        MoveJ speed 60 deg/s, acceleration 80 deg/s^2 (useActiveTCP=true optimoveEnabled=false optiMoveSpeed=0.3 optiMoveAcceleration=0.09) feature=Base
          Waypoint Waypoint_104: TCP in base x=-333.293 y=-480.744 z=350.142 mm, rx=2.2175 ry=0.1409 rz=2.2091 rad; joints [-82.414, -101.687, -97.87, -162.913, 4.302, 96.426] deg
        SuppressedNode
          Weight_value := get_weight()
    SuppressedNode
      Case (caseValue=38)
        SuppressedNode
          URCap VISOR Robotic App (SensoPart VISOR Robotic, SensoPart Industriesensorik GmbH) dataModel(visorAppTemplate=1); state(isChildrenLocked=true)
            URCap Easy Pick Setup (SensoPart VISOR Robotic, SensoPart Industriesensorik GmbH) dataModel(visorId=0, visorSetJob=true, visorJobName=Container_S_rack, visorImageAcqSetup=2, visorSetupStatus=2); state(isChildrenLocked=true)
            URCap Process (SensoPart VISOR Robotic, SensoPart Industriesensorik GmbH) dataModel(Variable(key=visorCounterVar, variable(name=easyPickCount_4, initializeExpression=0)), Variable(key=visorPartsFoundVar, variable(name=easyPickParts_4, initializeExpression=0))); state(isChildrenLocked=true)
              URCap Image Acquisition Pose (SensoPart VISOR Robotic, SensoPart Industriesensorik GmbH) state(isChildrenLocked=true)
              URCap Object Detected (SensoPart VISOR Robotic, SensoPart Industriesensorik GmbH) state(isChildrenLocked=true)
                Folder Open Gripper
                  Placeholder
                URCap Approach Pose (SensoPart VISOR Robotic, SensoPart Industriesensorik GmbH) state(isChildrenLocked=true)
                URCap Target Pose (SensoPart VISOR Robotic, SensoPart Industriesensorik GmbH) state(isChildrenLocked=true)
                Folder Close Gripper
                  Placeholder
                URCap Exit Pose (SensoPart VISOR Robotic, SensoPart Industriesensorik GmbH) state(isChildrenLocked=true)
              URCap No Object Detected (SensoPart VISOR Robotic, SensoPart Industriesensorik GmbH) dataModel(Variable(key=visorNoObjCountVar, variable(name=easyPickNoObj_4, initializeExpression=0)))
                Placeholder
    Case (caseValue=39)
      Folder Powder container Pick [hidden by the author, left out]
    Case (caseValue=40)
      Folder Decap Container  [hidden by the author, left out]
    Case (caseValue=41)
      Folder Place the open PowderA container & dosing
        SuppressedNode
          Script: tilt_to_home()
        SuppressedNode
          Script: tilt_send(4)
        URCap VISOR Robotic App (SensoPart VISOR Robotic, SensoPart Industriesensorik GmbH) dataModel(visorAppTemplate=1); state(isChildrenLocked=true)
          URCap Easy Pick Setup (SensoPart VISOR Robotic, SensoPart Industriesensorik GmbH) dataModel(visorId=0, visorImageAcqSetup=2, visorDetector=1, visorSetJob=true, visorOffsetSet=true, visorImageAcqSource=2, visorJobName=PoTS, visorSetupStatus=3, Pose(key=visorGripPose, Position(key=posePosition, Length(key=X value=-0.729991 unit=M), Length(key=Y value=-0.185228 unit=M), Length(key=Z value=0.248335 unit=M)), Rotation(key=poseRotation, Angle(key=RX value=-0.919003 unit=RAD), Angle(key=RY value=1.612625 unit=RAD), Angle(key=RZ value=-1.647622 unit=RAD))), Feature(key=visorImageAcqFeature name=Trigger)); state(isChildrenLocked=true)
          URCap Process (SensoPart VISOR Robotic, SensoPart Industriesensorik GmbH) dataModel(Variable(key=visorCounterVar, variable(name=easyPickCount_7, initializeExpression=0)), Variable(key=visorPartsFoundVar, variable(name=easyPickParts_7, initializeExpression=0))); state(isChildrenLocked=true)
            URCap Image Acquisition Pose (SensoPart VISOR Robotic, SensoPart Industriesensorik GmbH) state(isChildrenLocked=true)
            URCap Object Detected (SensoPart VISOR Robotic, SensoPart Industriesensorik GmbH) state(isChildrenLocked=true)
              Folder Open Gripper
                URCap Gripper (Robotiq_Grippers, Robotiq Inc.) dataModel(position=0.0, force=30.19607843137255, speed=30.19607843137255, positionInDouble=0.0, forceInDouble=30.19607843137255, speedInDouble=30.19607843137255, slaveIds=[9], blocking=true)
                SuppressedNode
                  Set NoAction tcp=TCP_fingers
                SuppressedNode
                  Wait Sleep waitTime=0.2
                MoveL speed 250 mm/s, acceleration 1200 mm/s^2 (useActiveTCP=true optimoveEnabled=false optiMoveSpeed=0.3 optiMoveAcceleration=0.09) feature=Base
                  Waypoint OP_PowderA2: TCP in base x=9.371 y=-409.434 z=294.169 mm, rx=-0.8233 ry=1.7094 rz=-1.6983 rad; joints [-57.265, -122.586, -76.992, -161.25, 72.295, 1.124] deg; TCP offset x=0 y=0 z=161 mm, rx=3.1415 ry=0 rz=0 rad
                  Waypoint OP_PowderA_ab_1: TCP in base x=-12.145 y=-363.335 z=315.326 mm, rx=-0.7771 ry=1.753 rz=-1.7409 rad; joints [-58.232, -116.012, -83.989, -160.83, 75.01, 1.147] deg; TCP offset x=0 y=0 z=161 mm, rx=3.1415 ry=0 rz=0 rad
                  Waypoint OP_PowderA_pick: TCP in base x=-19.99 y=-367.909 z=180.101 mm, rx=-0.5462 ry=1.936 rz=-1.9301 rad; joints [-66.516, -128.259, -85.768, -146.461, 83.267, 1.188] deg
                  URCap Gripper (Robotiq_Grippers, Robotiq Inc.) dataModel(position=100.0, force=30.19607843137255, speed=30.19607843137255, positionInDouble=100.0, forceInDouble=30.19607843137255, speedInDouble=30.19607843137255, slaveIds=[9], blocking=true)
                  Wait Sleep waitTime=0.5
                  Set DigitalOutput pin=GRP_3F_Open; digitalValue=1
                  SuppressedNode
                    Script: Motors_off()
                  Waypoint OP_PowderA_ab_2: motionParameters(jointSpeed=1.047198 jointAcceleration=1.396263 cartesianSpeed=0.05 cartesianAcceleration=0.3); TCP in base x=-12.145 y=-363.335 z=315.326 mm, rx=-0.7771 ry=1.753 rz=-1.7409 rad; joints [-58.232, -116.012, -83.989, -160.83, 75.01, 1.147] deg
                  Waypoint Op_PowA_wP: TCP in base x=-173.728 y=-372.934 z=295.117 mm, rx=-0.9724 ry=1.541 rz=-1.5487 rad; joints [-67.269, -106.894, -99.849, -153.52, 49.211, 1.028] deg
              URCap Approach Pose (SensoPart VISOR Robotic, SensoPart Industriesensorik GmbH) dataModel(visorOffsetZ=0.0, visorJointSpeed=25.0, visorJointAcc=30.0); state(isChildrenLocked=true)
              URCap Target Pose (SensoPart VISOR Robotic, SensoPart Industriesensorik GmbH) dataModel(visorToolSpeed=50.0, visorToolAcc=100.0); state(isChildrenLocked=true)
              Folder Close Gripper
                container_place := get_actual_tcp_pose()
                SuppressedNode
                  radius := 0.035
                SuppressedNode
                  PoTS_place_abov := pose_trans(container_place, p[0,0,radius,0,0,0])
                SuppressedNode
                  MoveL speed 50 mm/s, acceleration 500 mm/s^2 (useActiveTCP=true optimoveEnabled=false optiMoveSpeed=0.3 optiMoveAcceleration=0.09) feature=Base
                    Waypoint Variable (Variable): variable(name=PoTS_place_abov)
                target_pose := pose_trans(container_place, p[0,0.09,0,0,0,0])
                MoveL speed 50 mm/s, acceleration 500 mm/s^2 (useActiveTCP=true optimoveEnabled=false optiMoveSpeed=0.3 optiMoveAcceleration=0.09) feature=Base
                  Waypoint Variable (Variable): motionParameters(jointSpeed=1.047198 jointAcceleration=1.396263 cartesianSpeed=0.05 cartesianAcceleration=0.3); variable=target_pose
                URCap Gripper (Robotiq_Grippers, Robotiq Inc.) dataModel(position=0.0, force=30.19607843137255, speed=30.19607843137255, positionInDouble=0.0, forceInDouble=30.19607843137255, speedInDouble=30.19607843137255, slaveIds=[9], blocking=true)
              URCap Exit Pose (SensoPart VISOR Robotic, SensoPart Industriesensorik GmbH) dataModel(visorOffsetZ=-50.0); state(isChildrenLocked=true)
            URCap No Object Detected (SensoPart VISOR Robotic, SensoPart Industriesensorik GmbH) dataModel(Variable(key=visorNoObjCountVar, variable(name=easyPickNoObj_7, initializeExpression=0)))
              Popup Message (haltProgram=false message=No weigh scale detected inputType=Text)
        place_pose := get_actual_tcp_pose()
        Script: center_pose()
        SuppressedNode
          center_tilt_pos := P_center
        MoveJ speed 60 deg/s, acceleration 80 deg/s^2 (useActiveTCP=true optimoveEnabled=false optiMoveSpeed=0.3 optiMoveAcceleration=0.09) feature=Base
          Waypoint Waypoint_1: TCP in base x=-451.049 y=-340.589 z=308.224 mm, rx=0.0971 ry=0.091 rz=-1.5784 rad; joints [-127.334, -100.578, -80.109, -94.907, 86.186, -126.663] deg
    Case (caseValue=42)
      Folder Powder Emptying [hidden by the author, left out]
    Case (caseValue=43)
      Folder Powder dosing
        SuppressedNode
          Script: zero_scale()
        Script: send_target_info()
        Script: send_powder_info()
        switch_spat_M := True
        switch_spat_S := True
        switch_spat_F_S := True
        Timer (action=Start) variable(name=Dosing_time)
        SuppressedNode
          Script: tilt_to_home()
        SuppressedNode
          Folder spatula_selection test
            weight_value := get_weight()
            diff := target_weight-weight_value
            Script: scooping_init()
            Script: compute_level_percent(W_now, weight_value)
            Script: spatula = select_spatula(Pow_name, level, diff)
        URCap VISOR Robotic App (SensoPart VISOR Robotic, SensoPart Industriesensorik GmbH) dataModel(visorAppTemplate=1); state(isChildrenLocked=true)
          URCap Easy Pick Setup (SensoPart VISOR Robotic, SensoPart Industriesensorik GmbH) dataModel(visorId=0, visorSetJob=true, visorImageAcqSetup=2, visorCalibSetNo=9, visorDetector=1, visorImageAcqSource=2, visorJobName=Weight_scale, visorOffsetSet=true, visorSetupStatus=3, Pose(key=visorGripPose, Position(key=posePosition, Length(key=X value=-0.45122 unit=M), Length(key=Y value=0.110677 unit=M), Length(key=Z value=0.129785 unit=M)), Rotation(key=poseRotation, Angle(key=RX value=0.852924 unit=RAD), Angle(key=RY value=1.33496 unit=RAD), Angle(key=RZ value=-0.958582 unit=RAD))), Feature(key=visorImageAcqFeature name=Trigger)); state(isChildrenLocked=true)
          URCap Process (SensoPart VISOR Robotic, SensoPart Industriesensorik GmbH) dataModel(Variable(key=visorCounterVar, variable=easyPickCount_4), Variable(key=visorPartsFoundVar, variable=easyPickParts_4)); state(isChildrenLocked=true)
            URCap Image Acquisition Pose (SensoPart VISOR Robotic, SensoPart Industriesensorik GmbH) state(isChildrenLocked=true)
            URCap Object Detected (SensoPart VISOR Robotic, SensoPart Industriesensorik GmbH) state(isChildrenLocked=true)
              Folder Open Gripper
                Script: tare_scale()
                Wait Sleep waitTime=0.2
                weight_value := get_weight()
                Wait Sleep waitTime=0.2
                diff := target_weight-weight_value
                Script: scooping_init()
                Script: compute_level_percent(W_now, weight_value)
                Script: send_level_info()
                spatula := select_spatula(Pow_name, level, diff)
                SuppressedNode
                  spatula := select_spatula(Flowability,level,diff,density)
                SuppressedNode
                  Script: spatula = "spatula_M"
                Wait Sleep waitTime=0.2
                Script: send_spatula_info()
                If spatula ≟ "spatula_L"
                  MoveJ speed 60 deg/s, acceleration 80 deg/s^2 (useActiveTCP=true optimoveEnabled=false optiMoveSpeed=0.3 optiMoveAcceleration=0.09) feature=Base
                    Waypoint Spatula_otw: TCP in base x=-222.06 y=-318.141 z=425.288 mm, rx=-0.0004 ry=-0.0001 rz=3.0344 rad; joints [-104.723, -74.795, -88.594, -106.601, 90.132, -8.655] deg
                    Waypoint pick_spat_L_abv: TCP in base x=239.059 y=-67.213 z=280.721 mm, rx=0 ry=-0.0005 rz=3.1068 rad; joints [16.774, -49.077, -122.624, -98.282, 90.162, 108.776] deg
                  MoveL speed 250 mm/s, acceleration 1200 mm/s^2 (useActiveTCP=true optimoveEnabled=false optiMoveSpeed=0.3 optiMoveAcceleration=0.09) feature=Base
                    Waypoint spat_L_pick: TCP in base x=242.469 y=-67.302 z=193.171 mm, rx=0 ry=-0.0005 rz=3.1068 rad; joints [16.429, -49.275, -135.385, -85.324, 90.17, 108.483] deg
                    URCap Gripper (Robotiq_Grippers, Robotiq Inc.) dataModel(position=100.0, force=30.0, speed=0.0, positionInDouble=100.0, forceInDouble=30.0, speedInDouble=0.0, slaveIds=[9], blocking=true)
                    Waypoint spat_L_lift: motionParameters(blendRadius=0.01); TCP in base x=245.402 y=-67.432 z=289.049 mm, rx=0 ry=-0.0005 rz=3.1068 rad; joints [16.24, -50.411, -121.005, -98.568, 90.16, 108.238] deg
                    Waypoint spat_L_side: motionParameters(blendRadius=0.01); TCP in base x=247.134 y=-17.634 z=289.063 mm, rx=0 ry=-0.0005 rz=3.1068 rad; joints [28.487, -49.174, -121.365, -99.443, 90.16, 120.484] deg
                    Waypoint spat_L_up: motionParameters(blendRadius=0.05); TCP in base x=247.136 y=-17.665 z=397.131 mm, rx=0 ry=-0.0005 rz=3.1068 rad; joints [28.565, -53.55, -103.607, -112.824, 90.132, 120.503] deg
                  MoveJ speed 60 deg/s, acceleration 80 deg/s^2 (useActiveTCP=true optimoveEnabled=false optiMoveSpeed=0.3 optiMoveAcceleration=0.09) feature=Base
                    Waypoint Spatula_otw: TCP in base x=-222.06 y=-318.141 z=425.288 mm, rx=-0.0004 ry=-0.0001 rz=3.0344 rad; joints [-104.723, -74.795, -88.594, -106.601, 90.132, -8.655] deg
                ElseIf spatula ≟"spatula_M"
                  MoveJ speed 60 deg/s, acceleration 80 deg/s^2 (useActiveTCP=true optimoveEnabled=false optiMoveSpeed=0.3 optiMoveAcceleration=0.09) feature=Base
                    Waypoint Spatula_otw: TCP in base x=-222.06 y=-318.141 z=425.288 mm, rx=-0.0004 ry=-0.0001 rz=3.0344 rad; joints [-104.723, -74.795, -88.594, -106.601, 90.132, -8.655] deg
                    Waypoint spat_M_up: motionParameters(blendRadius=0.05); TCP in base x=245.496 y=-112.113 z=420.344 mm, rx=0 ry=-0.0005 rz=3.0677 rad; joints [5.167, -58.065, -98.393, -113.528, 90.127, 99.337] deg
                  MoveL speed 250 mm/s, acceleration 1200 mm/s^2 (useActiveTCP=true optimoveEnabled=false optiMoveSpeed=0.3 optiMoveAcceleration=0.09) feature=Base
                    Waypoint spat_M_pick: TCP in base x=244.674 y=-111.985 z=192.299 mm, rx=0 ry=-0.0005 rz=3.0677 rad; joints [5.062, -53.127, -134.29, -82.569, 90.166, 99.363] deg
                    URCap Gripper (Robotiq_Grippers, Robotiq Inc.) dataModel(position=100.0, force=30.0, speed=0.0, positionInDouble=100.0, forceInDouble=30.0, speedInDouble=0.0, slaveIds=[9], blocking=true)
                    Waypoint spat_M_up: motionParameters(blendRadius=0.05); TCP in base x=245.496 y=-112.113 z=420.344 mm, rx=0 ry=-0.0005 rz=3.0677 rad; joints [5.167, -58.065, -98.393, -113.528, 90.127, 99.337] deg
                    Waypoint Spatula_otw: TCP in base x=-222.06 y=-318.141 z=425.288 mm, rx=-0.0004 ry=-0.0001 rz=3.0344 rad; joints [-104.723, -74.795, -88.594, -106.601, 90.132, -8.655] deg
                  switch_spat_M := False
                ElseIf spatula≟"spatula_S"
                  MoveJ speed 60 deg/s, acceleration 80 deg/s^2 (useActiveTCP=true optimoveEnabled=false optiMoveSpeed=0.3 optiMoveAcceleration=0.09) feature=Base
                    Waypoint Spatula_otw: TCP in base x=-222.06 y=-318.141 z=425.288 mm, rx=-0.0004 ry=-0.0001 rz=3.0344 rad; joints [-104.723, -74.795, -88.594, -106.601, 90.132, -8.655] deg
                    Waypoint spat_S_Up_7: motionParameters(blendRadius=0.05); TCP in base x=252.088 y=-159.242 z=423.282 mm, rx=0 ry=-0.0005 rz=3.0677 rad; joints [-5.618, -62.24, -96.192, -111.556, 90.127, 88.551] deg
                  MoveL speed 250 mm/s, acceleration 1200 mm/s^2 (useActiveTCP=true optimoveEnabled=false optiMoveSpeed=0.3 optiMoveAcceleration=0.09) feature=Base
                    Waypoint spat_S_Pick_4: TCP in base x=245.377 y=-158.668 z=192.286 mm, rx=0 ry=-0.0005 rz=3.0677 rad; joints [-5.78, -57.937, -132.467, -79.585, 90.161, 88.525] deg
                    URCap Gripper (Robotiq_Grippers, Robotiq Inc.) dataModel(position=100.0, force=30.0, speed=0.0, positionInDouble=100.0, forceInDouble=30.0, speedInDouble=0.0, slaveIds=[9], blocking=true)
                    Waypoint spat_S_Up_8: motionParameters(blendRadius=0.05); TCP in base x=252.088 y=-159.242 z=423.282 mm, rx=0 ry=-0.0005 rz=3.0677 rad; joints [-5.618, -62.24, -96.192, -111.556, 90.127, 88.551] deg
                    Waypoint Spatula_otw: TCP in base x=-222.06 y=-318.141 z=425.288 mm, rx=-0.0004 ry=-0.0001 rz=3.0344 rad; joints [-104.723, -74.795, -88.594, -106.601, 90.132, -8.655] deg
                  switch_spat_S := False
                ElseIf spatula≟"spatula_flat_M"
                  MoveJ speed 60 deg/s, acceleration 80 deg/s^2 (useActiveTCP=true optimoveEnabled=false optiMoveSpeed=0.3 optiMoveAcceleration=0.09) feature=Base
                    Waypoint Spatula_otw: TCP in base x=-222.06 y=-318.141 z=425.288 mm, rx=-0.0004 ry=-0.0001 rz=3.0344 rad; joints [-104.723, -74.795, -88.594, -106.601, 90.132, -8.655] deg
                    Waypoint spat_flatM_up: motionParameters(blendRadius=0.05); TCP in base x=229.023 y=-211.443 z=418.634 mm, rx=0 ry=-0.0005 rz=3.0677 rad; joints [-17.294, -63.925, -96.117, -109.949, 90.128, 76.878] deg
                  MoveL speed 250 mm/s, acceleration 1200 mm/s^2 (useActiveTCP=true optimoveEnabled=false optiMoveSpeed=0.3 optiMoveAcceleration=0.09) feature=Base
                    Waypoint spat_flatM_pick: TCP in base x=241.029 y=-208.057 z=192.271 mm, rx=0 ry=-0.0005 rz=3.0677 rad; joints [-16.075, -63.047, -130.143, -76.801, 90.154, 78.231] deg
                    URCap Gripper (Robotiq_Grippers, Robotiq Inc.) dataModel(position=100.0, force=30.0, speed=0.0, positionInDouble=100.0, forceInDouble=30.0, speedInDouble=0.0, slaveIds=[9], blocking=true, robotCompliant=false)
                    Waypoint spat_flatM_up: motionParameters(blendRadius=0.05); TCP in base x=229.023 y=-211.443 z=418.634 mm, rx=0 ry=-0.0005 rz=3.0677 rad; joints [-17.294, -63.925, -96.117, -109.949, 90.128, 76.878] deg
                    Waypoint Spatula_otw: TCP in base x=-222.06 y=-318.141 z=425.288 mm, rx=-0.0004 ry=-0.0001 rz=3.0344 rad; joints [-104.723, -74.795, -88.594, -106.601, 90.132, -8.655] deg
                  switch_spat_F_M := False
                ElseIf spatula≟"spatula_flat_S"
                  MoveJ speed 60 deg/s, acceleration 80 deg/s^2 (useActiveTCP=true optimoveEnabled=false optiMoveSpeed=0.3 optiMoveAcceleration=0.09) feature=Base
                    Waypoint Spatula_otw: TCP in base x=-222.06 y=-318.141 z=425.288 mm, rx=-0.0004 ry=-0.0001 rz=3.0344 rad; joints [-104.723, -74.795, -88.594, -106.601, 90.132, -8.655] deg
                    Waypoint spat_flatS_up: motionParameters(blendRadius=0.05); TCP in base x=237.652 y=-253.944 z=403.961 mm, rx=0 ry=-0.0005 rz=3.0677 rad; joints [-24.273, -68.411, -95.947, -105.635, 90.132, 69.906] deg
                  MoveL speed 250 mm/s, acceleration 1200 mm/s^2 (useActiveTCP=true optimoveEnabled=false optiMoveSpeed=0.3 optiMoveAcceleration=0.09) feature=Base
                    Waypoint spat_flatS_pick: TCP in base x=241.326 y=-251.726 z=192.257 mm, rx=0 ry=-0.0005 rz=3.0677 rad; joints [-23.749, -68.568, -127.154, -74.27, 90.149, 70.556] deg
                    URCap Gripper (Robotiq_Grippers, Robotiq Inc.) dataModel(position=100.0, force=30.0, speed=0.0, positionInDouble=100.0, forceInDouble=30.0, speedInDouble=0.0, slaveIds=[9], blocking=true, robotCompliant=false)
                    Waypoint spat_flatS_up: motionParameters(blendRadius=0.05); TCP in base x=237.652 y=-253.944 z=403.961 mm, rx=0 ry=-0.0005 rz=3.0677 rad; joints [-24.273, -68.411, -95.947, -105.635, 90.132, 69.906] deg
                    Waypoint Spatula_otw: TCP in base x=-222.06 y=-318.141 z=425.288 mm, rx=-0.0004 ry=-0.0001 rz=3.0344 rad; joints [-104.723, -74.795, -88.594, -106.601, 90.132, -8.655] deg
                  switch_spat_F_S := False
                weight_value := get_weight()
                Script: auto_tilt_and_scoop(W_now, target_weight, weight_value)
              URCap Approach Pose (SensoPart VISOR Robotic, SensoPart Industriesensorik GmbH) dataModel(visorJointSpeed=10.0, visorJointAcc=15.0, visorOffsetZ=0.0); state(isChildrenLocked=true)
              URCap Target Pose (SensoPart VISOR Robotic, SensoPart Industriesensorik GmbH) dataModel(visorToolSpeed=20.0, visorToolAcc=50.0); state(isChildrenLocked=true)
              Folder Close Gripper
                dispense_pos := get_actual_tcp_pose()
                Loop While (checkContinuously=true) expression=weight_value≤target_weight
                  MoveL speed 250 mm/s, acceleration 1200 mm/s^2 (useActiveTCP=true optimoveEnabled=false optiMoveSpeed=0.3 optiMoveAcceleration=0.09) feature=Base
                    Waypoint Variable (Variable): motionParameters(jointSpeed=0.436332 jointAcceleration=0.523599 cartesianSpeed=0.1 cartesianAcceleration=0.2); variable=dispense_pos
                    Script: log_weight()
                    Wait Sleep waitTime=0.5
                    If level≥90.0
                      Script: Rotate()
                    If level≤85
                      Script: tilt_to_home()
                    Wait Sleep waitTime=0.5
                    Start_thread := True
                    vib_thread := True
                    SuppressedNode
                      tilt_angle := current_pose[5]
                    Wait Sleep waitTime=0.5
                    SuppressedNode
                      Loop While (checkContinuously=true) expression=diff>3.0
                        tilt_pose := pose_trans(get_actual_tcp_pose(), p[0, 0, 0, 0, 0, 1.0])
                        Script: movel(tilt_pose, a=0.1, v=0.1, r=0.00001)
                        tilt_pose := pose_trans(get_actual_tcp_pose(), p[0, 0, 0, 0, 0, -1.0])
                        Script: movel(tilt_pose, a=0.1, v=0.1, r=0.00001)
                    If diff ≥(target_g)
                      tilt_pose := pose_trans(get_actual_tcp_pose(), p[0, 0, 0, 0, 0, 2.0])
                      Script: movel(tilt_pose, a=0.1, v=0.1, r=0.00001)
                    Else 
                      Loop While (checkContinuously=true) expression=weight_value≤target_weight and tilt_angle≥(-1.999) and tilt_angle≤0.5
                        current_error := target_weight-weight_value
                        Integral_error := Integral_error+current_error*dt
                        derivative := (current_error-previous_error)/dt
                        tilt_increment := (kp*current_error)+(ki*Integral_error)+(kd*derivative)
                        current_pose := get_actual_tcp_pose()
                        tilt_angle := current_pose[5]
                        tilt_pose := pose_trans(current_pose, p[0, 0, 0, 0, 0, tilt_increment])
                        Script: movel(tilt_pose, a=0.1, v=0.1, r=0.00001)
                        previous_error := current_error
                    Start_thread := False
                    SuppressedNode
                      Waypoint Waypoint_64: motionParameters(jointSpeed=1.047198 jointAcceleration=1.396263 cartesianSpeed=0.03 cartesianAcceleration=0.1 blendRadius=0.05); TCP in base x=-542.998 y=-117.021 z=221.977 mm, rx=1.8981 ry=-0.7227 rz=1.5827 rad; joints [-123.845, -120.87, -101.018, -172.406, 14.907, 127.864] deg
                    weight_value := get_weight()
                    tilt_angle := -1
                    Wait Sleep waitTime=0.5
                    vib_thread := False
                    MoveL speed 250 mm/s, acceleration 500 mm/s^2 (useActiveTCP=true optimoveEnabled=false optiMoveSpeed=0.3 optiMoveAcceleration=0.09) feature=Base
                      Waypoint Variable (Variable): variable=dispense_pos
                    Script: compute_level_percent(W_now, weight_value)
                    Script: send_level_info()
                    Script: spatula = select_spatula(Pow_name, level, diff)
                    SuppressedNode
                      spatula := select_spatula(Flowability,level,diff,density)
                    SuppressedNode
                      Script: spatula = "spatula_M"
                    Wait Sleep waitTime=0.2
                    SuppressedNode
                      Script: spatula = str_cat("", spatula)
                    Integral_error := 0
                    current_error := 0
                    previous_error := 0
                    Set AnalogOutput pin=analog_out[0]; analogValue=0
                    Wait Sleep waitTime=0.2
                    Script: send_spatula_info()
                    If spatula ≟ "spatula_M" and switch_spat_M≟ True
                      MoveJ speed 60 deg/s, acceleration 80 deg/s^2 (useActiveTCP=true optimoveEnabled=false optiMoveSpeed=0.3 optiMoveAcceleration=0.09) feature=Base
                        Waypoint Spatula_otw: motionParameters(blendRadius=0.05); TCP in base x=-222.06 y=-318.141 z=425.288 mm, rx=-0.0004 ry=-0.0001 rz=3.0344 rad; joints [-104.723, -74.795, -88.594, -106.601, 90.132, -8.655] deg
                        Waypoint spat_L_up: TCP in base x=247.136 y=-17.665 z=397.131 mm, rx=0 ry=-0.0005 rz=3.1068 rad; joints [28.565, -53.55, -103.607, -112.824, 90.132, 120.503] deg
                      MoveL speed 250 mm/s, acceleration 1200 mm/s^2 (useActiveTCP=true optimoveEnabled=false optiMoveSpeed=0.3 optiMoveAcceleration=0.09) feature=Base
                        Waypoint spat_L_side: TCP in base x=247.134 y=-17.634 z=289.063 mm, rx=0 ry=-0.0005 rz=3.1068 rad; joints [28.487, -49.174, -121.365, -99.443, 90.16, 120.484] deg
                        Waypoint spat_L_lift: TCP in base x=245.402 y=-67.432 z=289.049 mm, rx=0 ry=-0.0005 rz=3.1068 rad; joints [16.24, -50.411, -121.005, -98.568, 90.16, 108.238] deg
                        Waypoint spat_L_pick: TCP in base x=242.469 y=-67.302 z=193.171 mm, rx=0 ry=-0.0005 rz=3.1068 rad; joints [16.429, -49.275, -135.385, -85.324, 90.17, 108.483] deg
                        URCap Gripper (Robotiq_Grippers, Robotiq Inc.) dataModel(position=0.0, force=30.0, speed=100.0, positionInDouble=0.0, forceInDouble=30.0, speedInDouble=100.0, slaveIds=[9], blocking=true)
                        Waypoint spat_M_pick: TCP in base x=244.674 y=-111.985 z=192.299 mm, rx=0 ry=-0.0005 rz=3.0677 rad; joints [5.062, -53.127, -134.29, -82.569, 90.166, 99.363] deg
                        URCap Gripper (Robotiq_Grippers, Robotiq Inc.) dataModel(position=100.0, force=30.0, speed=0.0, positionInDouble=100.0, forceInDouble=30.0, speedInDouble=0.0, slaveIds=[9], blocking=true)
                        Waypoint spat_M_up: TCP in base x=245.496 y=-112.113 z=420.344 mm, rx=0 ry=-0.0005 rz=3.0677 rad; joints [5.167, -58.065, -98.393, -113.528, 90.127, 99.337] deg
                        Waypoint Spatula_otw: TCP in base x=-222.06 y=-318.141 z=425.288 mm, rx=-0.0004 ry=-0.0001 rz=3.0344 rad; joints [-104.723, -74.795, -88.594, -106.601, 90.132, -8.655] deg
                      switch_spat_M := False
                    ElseIf spatula ≟ "spatula_S" and switch_spat_S ≟ True
                      MoveL speed 250 mm/s, acceleration 1200 mm/s^2 (useActiveTCP=true optimoveEnabled=false optiMoveSpeed=0.3 optiMoveAcceleration=0.09) feature=Base
                        Waypoint Spatula_otw: motionParameters(blendRadius=0.05); TCP in base x=-222.06 y=-318.141 z=425.288 mm, rx=-0.0004 ry=-0.0001 rz=3.0344 rad; joints [-104.723, -74.795, -88.594, -106.601, 90.132, -8.655] deg
                        Waypoint spat_M_up: TCP in base x=245.496 y=-112.113 z=420.344 mm, rx=0 ry=-0.0005 rz=3.0677 rad; joints [5.167, -58.065, -98.393, -113.528, 90.127, 99.337] deg
                        Waypoint spat_M_pick: TCP in base x=244.674 y=-111.985 z=192.299 mm, rx=0 ry=-0.0005 rz=3.0677 rad; joints [5.062, -53.127, -134.29, -82.569, 90.166, 99.363] deg
                        URCap Gripper (Robotiq_Grippers, Robotiq Inc.) dataModel(position=0.0, force=30.19607843137255, speed=100.0, positionInDouble=0.0, forceInDouble=30.19607843137255, speedInDouble=100.0, slaveIds=[9], blocking=true)
                        Waypoint spat_S_pick: TCP in base x=238.159 y=-157.927 z=192.632 mm, rx=0 ry=-0.0005 rz=3.0677 rad; joints [-5.778, -56.616, -132.95, -80.422, 90.162, 88.526] deg
                        URCap Gripper (Robotiq_Grippers, Robotiq Inc.) dataModel(position=100.0, force=30.19607843137255, speed=0.0, positionInDouble=100.0, forceInDouble=30.19607843137255, speedInDouble=0.0, slaveIds=[9], blocking=true)
                        Waypoint spat_S_up: TCP in base x=244.261 y=-164.467 z=417.088 mm, rx=0 ry=-0.0005 rz=3.0677 rad; joints [-6.934, -61.411, -97.537, -111.041, 90.129, 87.239] deg
                        Waypoint Spatula_otw: TCP in base x=-222.06 y=-318.141 z=425.288 mm, rx=-0.0004 ry=-0.0001 rz=3.0344 rad; joints [-104.723, -74.795, -88.594, -106.601, 90.132, -8.655] deg
                      switch_spat_S := False
                    ElseIf spatula≟"spatula_flat_S"  and switch_spat_F_S ≟ True
                      MoveL speed 250 mm/s, acceleration 1200 mm/s^2 (useActiveTCP=true optimoveEnabled=false optiMoveSpeed=0.3 optiMoveAcceleration=0.09) feature=Base
                        Waypoint Spatula_otw: motionParameters(blendRadius=0.05); TCP in base x=-222.06 y=-318.141 z=425.288 mm, rx=-0.0004 ry=-0.0001 rz=3.0344 rad; joints [-104.723, -74.795, -88.594, -106.601, 90.132, -8.655] deg
                        Waypoint spat_flatM_up: TCP in base x=229.023 y=-211.443 z=418.634 mm, rx=0 ry=-0.0005 rz=3.0677 rad; joints [-17.294, -63.925, -96.117, -109.949, 90.128, 76.878] deg
                        Waypoint spat_flatM_pick: TCP in base x=241.029 y=-208.057 z=192.271 mm, rx=0 ry=-0.0005 rz=3.0677 rad; joints [-16.075, -63.047, -130.143, -76.801, 90.154, 78.231] deg
                        URCap Gripper (Robotiq_Grippers, Robotiq Inc.) dataModel(position=0.0, force=30.0, speed=0.0, positionInDouble=0.0, forceInDouble=30.0, speedInDouble=0.0, slaveIds=[9], blocking=true, robotCompliant=false)
                        Waypoint spat_flatS_pick: TCP in base x=241.326 y=-251.726 z=192.257 mm, rx=0 ry=-0.0005 rz=3.0677 rad; joints [-23.749, -68.568, -127.154, -74.27, 90.149, 70.556] deg
                        URCap Gripper (Robotiq_Grippers, Robotiq Inc.) dataModel(position=100.0, force=30.0, speed=0.0, positionInDouble=100.0, forceInDouble=30.0, speedInDouble=0.0, slaveIds=[9], blocking=true, robotCompliant=false)
                        Waypoint spat_flatS_up: TCP in base x=237.652 y=-253.944 z=403.961 mm, rx=0 ry=-0.0005 rz=3.0677 rad; joints [-24.273, -68.411, -95.947, -105.635, 90.132, 69.906] deg
                        Waypoint Spatula_otw: TCP in base x=-222.06 y=-318.141 z=425.288 mm, rx=-0.0004 ry=-0.0001 rz=3.0344 rad; joints [-104.723, -74.795, -88.594, -106.601, 90.132, -8.655] deg
                      switch_spat_F_S := False
                    Script: auto_tilt_and_scoop(W_now, target_weight, weight_value)
                    Wait Sleep waitTime=0.5
                Start_thread := False
                Wait Sleep waitTime=0.5
                vib_thread := False
                SuppressedNode
                  Script: Rotate()
              URCap Exit Pose (SensoPart VISOR Robotic, SensoPart Industriesensorik GmbH) dataModel(visorOffsetZ=0.0); state(isChildrenLocked=true)
            URCap No Object Detected (SensoPart VISOR Robotic, SensoPart Industriesensorik GmbH) dataModel(Variable(key=visorNoObjCountVar, variable=easyPickNoObj_4))
              Popup Message (haltProgram=false message=No weigh scale detected inputType=Text)
        SuppressedNode
          Task := "Dosing"
        SuppressedNode
          Script: scooping_init()
        MoveJ speed 60 deg/s, acceleration 80 deg/s^2 (useActiveTCP=true optimoveEnabled=false optiMoveSpeed=0.3 optiMoveAcceleration=0.09) feature=Base
          Waypoint Variable (Variable): motionParameters(jointSpeed=0.436332 jointAcceleration=0.523599 cartesianSpeed=0.1 cartesianAcceleration=0.2); variable=dispense_pos
        Script: after_scoop()
        Timer (action=Stop) variable=Dosing_time
        Script: send_dosing_time(Dosing_time)
        Timer (action=Reset) variable=Dosing_time
        Script: Dosing_done()
        Folder Place the Spatula back in the holder [hidden by the author, left out]
        SuppressedNode
          Folder powder dispensing
            SuppressedNode
              Target_weight := Target_weight/1000
            Loop While (checkContinuously=false) expression=Weight_value<Target_weight
              Script: auto_tilt_and_scoop(W_now, Target_weight, Weight_value)
              Start_thread := True
              MoveL speed 250 mm/s, acceleration 1200 mm/s^2 (useActiveTCP=true optimoveEnabled=false optiMoveSpeed=0.3 optiMoveAcceleration=0.09) feature=Base
                Waypoint Variable (Variable): motionParameters(jointSpeed=0.436332 jointAcceleration=0.523599 cartesianSpeed=0.05 cartesianAcceleration=0.2); variable=dispense_pos
                Wait Sleep waitTime=0.5
                Script: Rotate()
                Wait Sleep waitTime=0.5
              MoveL speed 250 mm/s, acceleration 1200 mm/s^2 (useActiveTCP=true optimoveEnabled=false optiMoveSpeed=0.3 optiMoveAcceleration=0.09) feature=Base
                Start_thread := True
                vib_mot_thread := True
                tilt_angle := current_pose[5]
                Wait Sleep waitTime=0.5
                SuppressedNode
                  Loop While (checkContinuously=true) expression=diff>3.0
                    tilt_pose := pose_trans(get_actual_tcp_pose(), p[0, 0, 0, 0, 0, 1.0])
                    Script: movel(tilt_pose, a=0.1, v=0.1, r=0.00001)
                    tilt_pose := pose_trans(get_actual_tcp_pose(), p[0, 0, 0, 0, 0, -1.0])
                    Script: movel(tilt_pose, a=0.1, v=0.1, r=0.00001)
                If diff>3.0
                  tilt_pose := pose_trans(get_actual_tcp_pose(), p[0, 0, 0, 0, 0, 2.0])
                  Script: movel(tilt_pose, a=0.1, v=0.1, r=0.00001)
                ElseIf diff≤3.0
                  Loop While (checkContinuously=false) expression=Weight_value≤Target_weight and tilt_angle≥(-1.999) and tilt_angle≤0
                    current_error := Target_weight-Weight_value
                    Integral_error := Integral_error+current_error*dt
                    derivative := (current_error-previous_error)/dt
                    tilt_increment := (kp*current_error)+(ki*Integral_error)+(kd*derivative)
                    current_pose := get_actual_tcp_pose()
                    tilt_angle := current_pose[5]
                    tilt_pose := pose_trans(current_pose, p[0, 0, 0, 0, 0, tilt_increment])
                    Script: movel(tilt_pose, a=0.1, v=0.1, r=0.00001)
                    previous_error := current_error
                Start_thread := False
                SuppressedNode
                  Waypoint Waypoint_64: motionParameters(jointSpeed=1.047198 jointAcceleration=1.396263 cartesianSpeed=0.03 cartesianAcceleration=0.1 blendRadius=0.05); TCP in base x=-542.998 y=-117.021 z=221.977 mm, rx=1.8981 ry=-0.7227 rz=1.5827 rad; joints [-123.845, -120.87, -101.018, -172.406, 14.907, 127.864] deg
                Weight_value := get_weight()
                Wait Sleep waitTime=0.5
                tilt_angle := -1
                vib_mot_thread := False
                MoveL speed 50 mm/s, acceleration 300 mm/s^2 (useActiveTCP=true optimoveEnabled=false optiMoveSpeed=0.3 optiMoveAcceleration=0.09) feature=Base
                  Waypoint Variable (Variable): motionParameters(jointSpeed=0.436332 jointAcceleration=0.523599 cartesianSpeed=0.05 cartesianAcceleration=0.2); variable=dispense_pos
                Integral_error := 0
                current_error := 0
                previous_error := 0
                Set AnalogOutput pin=analog_out[0]; analogValue=0
              Script: movel(pose_trans(dispense_pos, p[-0.02,0,0,0,0,0]))
            SuppressedNode
              MoveL speed 250 mm/s, acceleration 1200 mm/s^2 (useActiveTCP=true optimoveEnabled=false optiMoveSpeed=0.3 optiMoveAcceleration=0.09) feature=Base
                Waypoint aftr_scoo3: motionParameters(jointSpeed=1.047198 jointAcceleration=1.396263 cartesianSpeed=0.1 cartesianAcceleration=0.3); TCP in base x=-289.76 y=-315.385 z=303.744 mm, rx=0.16 ry=1.6274 rz=-0.3449 rad; joints [-76.632, -96.313, -113.776, -155.476, 32.027, -78.1] deg
                Waypoint ftr_scoop2: motionParameters(jointSpeed=1.047198 jointAcceleration=1.396263 cartesianSpeed=0.1 cartesianAcceleration=0.4); TCP in base x=194.287 y=-495.78 z=282.072 mm, rx=-0.179 ry=1.6121 rz=-0.016 rad; joints [-34.133, -129.723, -68.393, -165.549, 50.138, -80.843] deg
                Waypoint aftr_scoop1: motionParameters(jointSpeed=1.047198 jointAcceleration=1.396263 cartesianSpeed=0.1 cartesianAcceleration=0.4); TCP in base x=138.504 y=-514.48 z=214.154 mm, rx=-0.1348 ry=1.5599 rz=-0.0592 rad; joints [-39.422, -130.004, -76.262, -153.157, 47.788, -83.41] deg
                Waypoint After_disp_3: motionParameters(jointSpeed=1.047198 jointAcceleration=1.396263 cartesianSpeed=0.1 cartesianAcceleration=0.4); TCP in base x=125.935 y=-585.611 z=299.546 mm, rx=0.9596 ry=-0.1344 rz=2.8807 rad; joints [-54.056, -115.535, -63.235, -120.118, 65.773, 48.319] deg
                Set AnalogOutput pin=analog_out[0]; analogValue=3
                Wait Sleep waitTime=2
                Set AnalogOutput pin=analog_out[0]; analogValue=0
                Waypoint aftr_scoop1: TCP in base x=138.504 y=-514.48 z=214.154 mm, rx=-0.1348 ry=1.5599 rz=-0.0592 rad; joints [-39.422, -130.004, -76.262, -153.157, 47.788, -83.41] deg
                Waypoint ftr_scoop2: motionParameters(jointSpeed=1.047198 jointAcceleration=1.396263 cartesianSpeed=0.1 cartesianAcceleration=0.4); TCP in base x=194.287 y=-495.78 z=282.072 mm, rx=-0.179 ry=1.6121 rz=-0.016 rad; joints [-34.133, -129.723, -68.393, -165.549, 50.138, -80.843] deg
                Waypoint Waypoint_63: motionParameters(blendRadius=0.05); TCP in base x=101.295 y=-465.376 z=381.756 mm, rx=0.9726 ry=-0.1584 rz=2.8872 rad; joints [-48.863, -99.659, -71.872, -130.079, 68.56, 52.636] deg; TCP offset x=0 y=0 z=161 mm, rx=3.1415 ry=0 rz=0 rad
                Waypoint Start: motionParameters(jointSpeed=1.047198 jointAcceleration=1.396263 cartesianSpeed=0.15 cartesianAcceleration=0.6); TCP in base x=-33.065 y=-365.399 z=389.873 mm, rx=0 ry=0 rz=2.7258 rad; joints [-73.774, -70.638, -96.716, -102.629, 90.121, 40.001] deg; TCP offset x=0 y=0 z=161 mm, rx=3.1415 ry=0 rz=0 rad
                Popup Message (haltProgram=false message=Powder dispensed successfully... inputType=Text)
            SuppressedNode
              Script: tilt()
        SuppressedNode
          Script: tilt_send()
    Case (caseValue=44)
      Folder Decap Container for recipe [hidden by the author, left out]
    Case (caseValue=45)
      Folder Place the decapped container- recipe [hidden by the author, left out]
    Case (caseValue=46)
      Folder Powder dosing for recipe [hidden by the author, left out]
    Case (caseValue=47)
      Folder Pick containers [hidden by the author, left out]
    Case (caseValue=48)
      Folder QR detections [hidden by the author, left out]
    SuppressedNode
      Case (caseValue=49)
        Folder QR Parameterization
          Device_ID := 1
          MoveJ speed 60 deg/s, acceleration 80 deg/s^2 (useActiveTCP=true optimoveEnabled=false optiMoveSpeed=0.3 optiMoveAcceleration=0.09) feature=Base
            Waypoint Variable (Variable): variable(featureName=Position1)
          URCap VISOR Trigger (SensoPart VISOR Robotic, SensoPart Industriesensorik GmbH) dataModel(visorId=0, visorSetJob=true, visorJobName=QR detection, visorImageAcqSetup=1); state(isChildrenLocked=true)
          pos1_powder := visor_getResponse(Device_ID)
          Script: pos1_powder = extract_powder_name(pos1_powder)
          MoveJ speed 60 deg/s, acceleration 80 deg/s^2 (useActiveTCP=true optimoveEnabled=false optiMoveSpeed=0.3 optiMoveAcceleration=0.09) feature=Base
            Waypoint Variable (Variable): variable(featureName=Position2)
          URCap VISOR Trigger (SensoPart VISOR Robotic, SensoPart Industriesensorik GmbH) dataModel(visorId=0, visorSetJob=true, visorJobName=QR detection, visorImageAcqSetup=1); state(isChildrenLocked=true)
          pos2_powder := visor_getResponse(Device_ID)
          Script: pos2_powder = extract_powder_name(pos2_powder)
          MoveJ speed 60 deg/s, acceleration 80 deg/s^2 (useActiveTCP=true optimoveEnabled=false optiMoveSpeed=0.3 optiMoveAcceleration=0.09) feature=Base
            Waypoint Variable (Variable): variable(featureName=Position3)
          URCap VISOR Trigger (SensoPart VISOR Robotic, SensoPart Industriesensorik GmbH) dataModel(visorId=0, visorSetJob=true, visorJobName=QR detection, visorImageAcqSetup=1); state(isChildrenLocked=true)
          pos3_powder := visor_getResponse(Device_ID)
          Script: pos3_powder = extract_powder_name(pos3_powder)
  '=========='
  Folder PostSettings [hidden by the author, left out]
  SuppressedNode
    Switch expression=Action
      Case (caseValue=1)
        Folder Pick [hidden by the author, left out]
      Case (caseValue=2)
        Folder Place [hidden by the author, left out]
      Case (caseValue=3)
        Folder Push
          Action_Info := "push"
      Case (caseValue=4)
        Folder Pull
          Action_Info := "pull"
      SuppressedNode
        Case (caseValue=5)
          Placeholder
      Case (caseValue=6)
        Folder Drop the cap [hidden by the author, left out]
      Case (caseValue=7)
        Folder Load [hidden by the author, left out]
      Case (caseValue=8)
        Folder Unload [hidden by the author, left out]
      Case (caseValue=11)
        SuppressedNode
          Folder Place without opening gripper
            Action_Info := "place object without gripper opening"
            SuppressedNode
              Script: do_transition(pose_trans(FRM_Reference, PSE_T), keep_rxry=OBJ_Picked)
            Script: movel(FRM_Container_S, a=0.025, v=0.015, r=0.00001)
            Folder EXTT
              Switch expression=JIG
                Case (caseValue=1)
                  Folder 3FG
                    If OBJ_Picked
                      Set DigitalOutput pin=GRP_3F_Open; digitalValue=1
            If PSE_A_H≠PSE_Z
              If JNT_Q≠JNT_Z
                Script: movej(get_inverse_kin(pose_trans(FRM_Reference, PSE_A_H), qnear=JNT_Q), r=0.050)
              Else 
                Script: movej(pose_trans(FRM_Reference, PSE_A_H), r=0.050)
            If PSE_A≠PSE_Z
              If JNT_Q≠JNT_Z
                Script: movej(get_inverse_kin(pose_trans(FRM_Reference, PSE_A), qnear=JNT_Q), r=0.020)
              Else 
                Script: movej(pose_trans(FRM_Reference, PSE_A), r=0.020)
            MoveL speed 400 mm/s, acceleration 500 mm/s^2 (useActiveTCP=true optimoveEnabled=false optiMoveSpeed=0.3 optiMoveAcceleration=0.09) feature=FRM_Reference
              If PSE_T_H≠PSE_Z
                Waypoint Variable (Variable): motionParameters(blendRadius=0.01); variable=PSE_T_H
              Waypoint Variable (Variable): motionParameters(jointSpeed=1.047198 jointAcceleration=1.396263 cartesianSpeed=0.09 cartesianAcceleration=0.05); variable=PSE_T
                Until TOOL_CONTACT_DETECTION (allowActions=false retraction=NONE decelerationAcceleration=0.5 decelerationAngularAcceleration=34.906585)
              Force Frame feature=FRM_Reference; selection=[1, 1, 1, 0, 0, 0]; wrench=[0, 0, 0, 0, 0, 0]; limitsForce=[0.1, 0.1, 0.01, 1.047198, 1.047198, 1.047198]; limitsMotion=[0.1, 0.1, 0.1, 0.349066, 0.349066, 0.349066]
                Waypoint Variable (Variable): motionParameters(jointSpeed=1.047198 jointAcceleration=1.396263 cartesianSpeed=0.07 cartesianAcceleration=0.04); variable=PSE_T
              Folder EXTT
                Switch expression=JIG
                  Case (caseValue=1)
                    Folder 3FG
                      If OBJ_Picked
                        Set DigitalOutput pin=GRP_3F_Open; digitalValue=0
                        Wait Sleep waitTime=0.2
              Folder EOAT
                ''
      Case (caseValue=12)
        Folder Decap [hidden by the author, left out]
      Case (caseValue=13)
        Timer (action=Reset) variable=TMR_Barcode
        Folder Read [hidden by the author, left out]
      Case (caseValue=15)
        Folder Detect
          Action_Info := "detect"
      Case (caseValue=30)
        Folder Shake [hidden by the author, left out]
      Case (caseValue=31)
        Action_Info := "Pick_Vial"
        Folder Pick_Vial [hidden by the author, left out]
      Case (caseValue=32)
        SuppressedNode
          decap := False
        Folder decap_Vial [hidden by the author, left out]
      Case (caseValue=33)
        Folder Shake and liquid transfer [hidden by the author, left out]
      SuppressedNode
        Case (caseValue=34)
          SafeHome (positionOptionType=SPEED_AND_ACCELERATION speed=1.047198 acceleration=1.396263 nextMotionTime=2)
          MoveJ speed 60 deg/s, acceleration 80 deg/s^2 (useActiveTCP=true optimoveEnabled=false optiMoveSpeed=0.3 optiMoveAcceleration=0.09) feature=Base
            Waypoint Waypoint_93: motionParameters(jointSpeed=0.436332 jointAcceleration=0.523599 cartesianSpeed=0.25 cartesianAcceleration=1.2); TCP in base x=206.301 y=-401.796 z=209.941 mm, rx=0 ry=0 rz=1.5608 rad; joints [-45.627, -84.145, -113.025, -72.821, 90.127, -225.014] deg
          MoveL speed 250 mm/s, acceleration 1200 mm/s^2 (useActiveTCP=true optimoveEnabled=false optiMoveSpeed=0.3 optiMoveAcceleration=0.09) feature=Base
            Waypoint Waypoint_94: motionParameters(jointSpeed=1.047198 jointAcceleration=1.396263 cartesianSpeed=0.1 cartesianAcceleration=0.5); TCP in base x=200.866 y=-400.818 z=105.073 mm, rx=0 ry=0 rz=1.5608 rad; joints [-46.083, -90.669, -123.933, -55.389, 90.105, -225.416] deg
          URCap Gripper (Robotiq_Grippers, Robotiq Inc.) dataModel(position=100.0, force=27.84313725490196, speed=32.15686274509804, positionInDouble=100.0, forceInDouble=27.84313725490196, speedInDouble=32.15686274509804, slaveIds=[9], blocking=true)
          Wait Sleep waitTime=1
          MoveL speed 250 mm/s, acceleration 1200 mm/s^2 (useActiveTCP=true optimoveEnabled=false optiMoveSpeed=0.3 optiMoveAcceleration=0.09) feature=Base
            Waypoint Waypoint_95: motionParameters(jointSpeed=1.047198 jointAcceleration=1.396263 cartesianSpeed=0.1 cartesianAcceleration=0.5 blendRadius=0.05); TCP in base x=200.866 y=-400.818 z=325.177 mm, rx=0 ry=0 rz=1.5608 rad; joints [-46.018, -81.306, -98.396, -90.289, 90.129, -225.47] deg
          MoveJ speed 60 deg/s, acceleration 80 deg/s^2 (useActiveTCP=true optimoveEnabled=false optiMoveSpeed=0.3 optiMoveAcceleration=0.09) feature=Base
            Waypoint Waypoint_96: motionParameters(jointSpeed=0.436332 jointAcceleration=0.523599 cartesianSpeed=0.25 cartesianAcceleration=1.2 blendRadius=0.05); TCP in base x=-615.829 y=233.809 z=300 mm, rx=0.0051 ry=0.0087 rz=-2.1118 rad; joints [-188.832, -110.936, -69.076, -89.912, 89.674, -157.919] deg
          MoveL speed 250 mm/s, acceleration 1200 mm/s^2 (useActiveTCP=true optimoveEnabled=false optiMoveSpeed=0.3 optiMoveAcceleration=0.09) feature=Base
            Waypoint Waypoint_97: motionParameters(jointSpeed=1.047198 jointAcceleration=1.396263 cartesianSpeed=0.1 cartesianAcceleration=0.5); TCP in base x=-615.829 y=233.809 z=13.91 mm, rx=0.0051 ry=0.0087 rz=-2.1118 rad; joints [-188.874, -123.68, -94.539, -51.707, 89.657, -157.833] deg
          URCap Gripper (Robotiq_Grippers, Robotiq Inc.) dataModel(position=0.0, force=27.84313725490196, speed=32.15686274509804, positionInDouble=0.0, forceInDouble=27.84313725490196, speedInDouble=32.15686274509804, slaveIds=[9], blocking=true)
          MoveJ speed 60 deg/s, acceleration 80 deg/s^2 (useActiveTCP=true optimoveEnabled=false optiMoveSpeed=0.3 optiMoveAcceleration=0.09) feature=Base
            Waypoint Waypoint_98: motionParameters(jointSpeed=0.436332 jointAcceleration=0.523599 cartesianSpeed=0.25 cartesianAcceleration=1.2); TCP in base x=-615.829 y=233.809 z=300 mm, rx=0.0051 ry=0.0087 rz=-2.1118 rad; joints [-188.832, -110.936, -69.076, -89.912, 89.674, -157.919] deg
          SafeHome (positionOptionType=SPEED_AND_ACCELERATION speed=1.047198 acceleration=1.396263 nextMotionTime=2)
          SuppressedNode
            Folder Decap
              Action_Info := "decapping"
              Set DigitalOutput pin=GRP_3F_Enable; digitalValue=1
              Set DigitalOutput pin=GRP_3F_Decap; digitalValue=1
              Force Frame feature=Base; selection=[0, 0, 1, 0, 0, 0]; wrench=[0, 0, 1, 0, 0, 0]; limitsForce=[0.15, 0.15, 0.001, 1.047198, 1.047198, 1.047198]; limitsMotion=[0.1, 0.1, 0.1, 0.349066, 0.349066, 0.349066]
                Script: check_decapping(offset=0.015, timeout=10, abort=CMD_Hold)
              Set DigitalOutput pin=GRP_3F_Decap; digitalValue=0
              Set DigitalOutput pin=GRP_3F_Enable; digitalValue=0
              MoveL speed 250 mm/s, acceleration 1200 mm/s^2 (useActiveTCP=true optimoveEnabled=false optiMoveSpeed=0.3 optiMoveAcceleration=0.09) feature=Base
                Waypoint Waypoint_5: motionParameters(jointSpeed=1.047198 jointAcceleration=1.396263 cartesianSpeed=0.1 cartesianAcceleration=0.5 blendRadius=0.05); TCP in base x=-31.859 y=-349.402 z=312.809 mm, rx=0 ry=0 rz=0 rad; joints [-72.832, -66.838, -110.376, -92.778, 90.139, -162.834] deg
              MoveJ speed 60 deg/s, acceleration 80 deg/s^2 (useActiveTCP=true optimoveEnabled=false optiMoveSpeed=0.3 optiMoveAcceleration=0.09) feature=Base
                Waypoint cap_dump: motionParameters(jointSpeed=0.436332 jointAcceleration=0.523599 cartesianSpeed=0.25 cartesianAcceleration=1.2); TCP in base x=-139.169 y=-420.164 z=146.096 mm, rx=0 ry=0 rz=0 rad; joints [-90.79, -86.479, -121, -62.513, 90.12, -180.712] deg
              URCap Gripper (Robotiq_Grippers, Robotiq Inc.) dataModel(position=0.0, force=100.0, speed=100.0, positionInDouble=0.0, forceInDouble=100.0, speedInDouble=100.0, slaveIds=[9], blocking=true)
              MoveJ speed 60 deg/s, acceleration 80 deg/s^2 (useActiveTCP=true optimoveEnabled=false optiMoveSpeed=0.3 optiMoveAcceleration=0.09) feature=Base
                Waypoint Waypoint_5: motionParameters(jointSpeed=0.436332 jointAcceleration=0.523599 cartesianSpeed=0.25 cartesianAcceleration=1.2 blendRadius=0.05); TCP in base x=-31.859 y=-349.402 z=312.809 mm, rx=0 ry=0 rz=0 rad; joints [-72.832, -66.838, -110.376, -92.778, 90.139, -162.834] deg
              Set DigitalOutput pin=digital_out[5]; digitalValue=1
      SuppressedNode
        Case (caseValue=35)
          Folder Pick the powder container
            URCap VISOR Robotic App (SensoPart VISOR Robotic, SensoPart Industriesensorik GmbH) dataModel(visorAppTemplate=1); state(isChildrenLocked=true)
              URCap Easy Pick Setup (SensoPart VISOR Robotic, SensoPart Industriesensorik GmbH) dataModel(visorId=0, visorSetJob=true, visorJobName=Container_S, visorImageAcqSetup=2, visorCalibSetNo=7, visorDetector=1, visorImageAcqSource=1, visorOffsetSet=true, visorSetupStatus=3, Pose(key=visorImageAcqPose, Position(key=posePosition, Length(key=X value=-0.51041 unit=M), Length(key=Y value=0.417301 unit=M), Length(key=Z value=0.464095 unit=M)), Rotation(key=poseRotation, Angle(key=RX value=0.000026 unit=RAD), Angle(key=RY value=-0.000024 unit=RAD), Angle(key=RZ value=-2.896187 unit=RAD))), Pose(key=visorGripPose, Position(key=posePosition, Length(key=X value=-0.52891 unit=M), Length(key=Y value=0.461593 unit=M), Length(key=Z value=-0.178186 unit=M)), Rotation(key=poseRotation, Angle(key=RX value=-0.279814 unit=RAD), Angle(key=RY value=2.118244 unit=RAD), Angle(key=RZ value=-2.110314 unit=RAD)))); state(isChildrenLocked=true)
              URCap Process (SensoPart VISOR Robotic, SensoPart Industriesensorik GmbH) dataModel(Variable(key=visorCounterVar, variable=easyPickCount), Variable(key=visorPartsFoundVar, variable=easyPickParts)); state(isChildrenLocked=true)
                URCap Image Acquisition Pose (SensoPart VISOR Robotic, SensoPart Industriesensorik GmbH) state(isChildrenLocked=true)
                URCap Object Detected (SensoPart VISOR Robotic, SensoPart Industriesensorik GmbH) state(isChildrenLocked=true)
                  Folder Open Gripper
                    URCap Gripper (Robotiq_Grippers, Robotiq Inc.) dataModel(position=0.0, force=30.0, speed=40.0, positionInDouble=0.0, forceInDouble=30.0, speedInDouble=40.0, slaveIds=[9], blocking=true)
                    MoveJ speed 60 deg/s, acceleration 80 deg/s^2 (useActiveTCP=true optimoveEnabled=false optiMoveSpeed=0.3 optiMoveAcceleration=0.09) feature=Base
                      Waypoint Waypoint_13: TCP in base x=-479.451 y=284.141 z=125.27 mm, rx=-0.2768 ry=2.0984 rz=-2.1213 rad; joints [-165.671, -112.009, -127.874, -95.426, 1.192, -23.029] deg
                  URCap Approach Pose (SensoPart VISOR Robotic, SensoPart Industriesensorik GmbH) dataModel(visorOffsetZ=-50.0); state(isChildrenLocked=true)
                  URCap Target Pose (SensoPart VISOR Robotic, SensoPart Industriesensorik GmbH) state(isChildrenLocked=true)
                  Folder Close Gripper
                    URCap Gripper (Robotiq_Grippers, Robotiq Inc.) dataModel(position=100.0, force=30.19607843137255, speed=40.0, positionInDouble=100.0, forceInDouble=30.19607843137255, speedInDouble=40.0, slaveIds=[9], blocking=true)
                  URCap Exit Pose (SensoPart VISOR Robotic, SensoPart Industriesensorik GmbH) dataModel(visorOffsetZ=-50.0); state(isChildrenLocked=true)
                URCap No Object Detected (SensoPart VISOR Robotic, SensoPart Industriesensorik GmbH) dataModel(Variable(key=visorNoObjCountVar, variable=easyPickNoObj))
                  Popup Message (haltProgram=false message=No Container detected inputType=Text)
            MoveJ speed 60 deg/s, acceleration 80 deg/s^2 (useActiveTCP=true optimoveEnabled=false optiMoveSpeed=0.3 optiMoveAcceleration=0.09) feature=Base
              SuppressedNode
                Waypoint Cont_midwa_1: motionParameters(jointSpeed=1.047198 jointAcceleration=1.396263 cartesianSpeed=0.25 cartesianAcceleration=1.2 blendRadius=0.01); TCP in base x=-462.252 y=294.856 z=204.322 mm, rx=-0.3472 ry=2.0343 rz=-2.0655 rad; joints [-166.773, -128.859, -129.893, 70.604, 5.32, -171.145] deg
              Waypoint Waypoint_70: motionParameters(jointSpeed=0.523599 jointAcceleration=0.698132 cartesianSpeed=0.25 cartesianAcceleration=1.2 blendRadius=0); TCP in base x=-472.821 y=292.44 z=207.418 mm, rx=-0.2598 ry=-2.0535 rz=2.0707 rad; joints [-170.164, -118.699, -96.461, -142.976, 25.725, -0.32] deg
              Waypoint Waypoint_78: motionParameters(jointSpeed=0.523599 jointAcceleration=0.872665 cartesianSpeed=0.25 cartesianAcceleration=1.2 blendRadius=0.05); TCP in base x=-51.45 y=-519.556 z=365.719 mm, rx=-1.2873 ry=1.0776 rz=-1.2185 rad; joints [-52.794, -108.287, -85.596, -162.721, 32.001, 1.948] deg
              Waypoint Waypoint_99: motionParameters(jointSpeed=0.523599 jointAcceleration=0.698132 cartesianSpeed=0.25 cartesianAcceleration=1.2 blendRadius=0.05); TCP in base x=-113.75 y=-390.11 z=317.307 mm, rx=-0.5194 ry=-0.8399 rz=1.7569 rad; joints [-108.345, -98.585, -86.606, -121.699, 124.957, 41.411] deg
            MoveL speed 250 mm/s, acceleration 1200 mm/s^2 (useActiveTCP=true optimoveEnabled=false optiMoveSpeed=0.3 optiMoveAcceleration=0.09) feature=Base
              Waypoint Waypoint_15: motionParameters(jointSpeed=1.047198 jointAcceleration=1.396263 cartesianSpeed=0.1 cartesianAcceleration=0.5 blendRadius=0.05); TCP in base x=29.144 y=-436.802 z=327.885 mm, rx=-0.5216 ry=-0.6236 rz=1.8627 rad; joints [-89.657, -89.204, -96.411, -97.086, 128.129, 64.023] deg
              Waypoint Waypoint_14: motionParameters(jointSpeed=1.047198 jointAcceleration=1.396263 cartesianSpeed=0.1 cartesianAcceleration=0.3); TCP in base x=68.712 y=-569.42 z=285.215 mm, rx=-0.6792 ry=-0.7121 rz=1.394 rad; joints [-90.137, -103.3, -96.148, -70.007, 141.633, 93.932] deg
              Waypoint Waypoint_100: motionParameters(jointSpeed=1.047198 jointAcceleration=1.396263 cartesianSpeed=0.05 cartesianAcceleration=0.3); TCP in base x=-47.22 y=-557.625 z=136.371 mm, rx=-0.6792 ry=-0.7121 rz=1.394 rad; joints [-101.643, -114.727, -100.71, -68.127, 140.302, 75.797] deg
            URCap Gripper (Robotiq_Grippers, Robotiq Inc.) dataModel(position=0.0, force=30.0, speed=40.0, positionInDouble=0.0, forceInDouble=30.0, speedInDouble=40.0, slaveIds=[9], blocking=true)
            MoveL speed 250 mm/s, acceleration 1200 mm/s^2 (useActiveTCP=true optimoveEnabled=false optiMoveSpeed=0.3 optiMoveAcceleration=0.09) feature=Base
              Waypoint Waypoint_25: motionParameters(jointSpeed=1.047198 jointAcceleration=1.396263 cartesianSpeed=0.1 cartesianAcceleration=0.3); TCP in base x=65.436 y=-569.388 z=287.821 mm, rx=-0.6792 ry=-0.7121 rz=1.394 rad; joints [-90.466, -103.248, -95.699, -70.925, 141.635, 93.398] deg
              Waypoint Waypoint_15: motionParameters(jointSpeed=1.047198 jointAcceleration=1.396263 cartesianSpeed=0.1 cartesianAcceleration=0.5 blendRadius=0.05); TCP in base x=29.144 y=-436.802 z=327.885 mm, rx=-0.5216 ry=-0.6236 rz=1.8627 rad; joints [-89.657, -89.204, -96.411, -97.086, 128.129, 64.023] deg
            SafeHome (positionOptionType=SPEED_AND_ACCELERATION speed=1.047198 acceleration=1.396263 nextMotionTime=2)
            SafeHome (positionOptionType=SPEED_AND_ACCELERATION speed=1.047198 acceleration=1.396263 nextMotionTime=2)
            SuppressedNode
              MoveJ speed 60 deg/s, acceleration 80 deg/s^2 (useActiveTCP=true optimoveEnabled=false optiMoveSpeed=0.3 optiMoveAcceleration=0.09) feature=Base
                Waypoint Container_midwa: motionParameters(blendRadius=0.05); TCP in base x=-379.239 y=-127.191 z=300 mm, rx=0 ry=0 rz=-1.2472 rad; joints [-141.945, -74.312, -107.466, -88.214, 90.137, -160.485] deg
            SuppressedNode
              URCap VISOR Robotic App (SensoPart VISOR Robotic, SensoPart Industriesensorik GmbH) dataModel(visorAppTemplate=1); state(isChildrenLocked=true)
                URCap Easy Pick Setup (SensoPart VISOR Robotic, SensoPart Industriesensorik GmbH) dataModel(visorId=0, visorSetJob=true, visorJobName=Target_container, visorImageAcqSetup=2, visorCalibSetNo=7, visorImageAcqSource=0, visorDetector=1, visorOffsetSet=true, visorSetupStatus=3, Pose(key=visorGripPose, Position(key=posePosition, Length(key=X value=-0.43018 unit=M), Length(key=Y value=0.500077 unit=M), Length(key=Z value=-0.155571 unit=M)), Rotation(key=poseRotation, Angle(key=RX value=0.000011 unit=RAD), Angle(key=RY value=0.000015 unit=RAD), Angle(key=RZ value=-2.896111 unit=RAD))), Pose(key=visorImageAcqPose, Position(key=posePosition, Length(key=X value=-0.391157 unit=M), Length(key=Y value=0.420635 unit=M), Length(key=Z value=0.411587 unit=M)), Rotation(key=poseRotation, Angle(key=RX value=-0.000006 unit=RAD), Angle(key=RY value=-0.000024 unit=RAD), Angle(key=RZ value=-2.896146 unit=RAD)))); state(isChildrenLocked=true)
                URCap Process (SensoPart VISOR Robotic, SensoPart Industriesensorik GmbH) dataModel(Variable(key=visorCounterVar, variable=easyPickCount_1), Variable(key=visorPartsFoundVar, variable=easyPickParts_1)); state(isChildrenLocked=true)
                  URCap Image Acquisition Pose (SensoPart VISOR Robotic, SensoPart Industriesensorik GmbH) state(isChildrenLocked=true)
                  URCap Object Detected (SensoPart VISOR Robotic, SensoPart Industriesensorik GmbH) state(isChildrenLocked=true)
                    Folder Open Gripper
                      URCap Gripper (Robotiq_Grippers, Robotiq Inc.) dataModel(position=0.0, force=30.0, speed=40.0, positionInDouble=0.0, forceInDouble=30.0, speedInDouble=40.0, slaveIds=[9], blocking=true)
                    URCap Approach Pose (SensoPart VISOR Robotic, SensoPart Industriesensorik GmbH) dataModel(visorOffsetZ=-50.0); state(isChildrenLocked=true)
                    URCap Target Pose (SensoPart VISOR Robotic, SensoPart Industriesensorik GmbH) state(isChildrenLocked=true)
                    Folder Close Gripper
                      URCap Gripper (Robotiq_Grippers, Robotiq Inc.) dataModel(position=100.0, force=30.19607843137255, speed=40.0, positionInDouble=100.0, forceInDouble=30.19607843137255, speedInDouble=40.0, slaveIds=[9], blocking=true)
                    URCap Exit Pose (SensoPart VISOR Robotic, SensoPart Industriesensorik GmbH) dataModel(visorOffsetZ=-50.0); state(isChildrenLocked=true)
                  URCap No Object Detected (SensoPart VISOR Robotic, SensoPart Industriesensorik GmbH) dataModel(Variable(key=visorNoObjCountVar, variable=easyPickNoObj_1))
                    Popup Message (haltProgram=false message=No Target container is detected inputType=Text)
            SuppressedNode
              MoveJ speed 60 deg/s, acceleration 80 deg/s^2 (useActiveTCP=true optimoveEnabled=false optiMoveSpeed=0.3 optiMoveAcceleration=0.09) feature=Base
                Waypoint Waypoint_16: motionParameters(jointSpeed=0.698132 jointAcceleration=0.872665 cartesianSpeed=0.25 cartesianAcceleration=1.2); TCP in base x=-389.004 y=141.378 z=266.753 mm, rx=0.0001 ry=-0.0001 rz=-2.8961 rad; joints [-181.152, -76.776, -110.541, -82.676, 90.144, -105.201] deg
                Waypoint Waypoint_17: motionParameters(jointSpeed=0.698132 jointAcceleration=0.872665 cartesianSpeed=0.25 cartesianAcceleration=1.2); TCP in base x=-35.034 y=-360.271 z=346.67 mm, rx=0.0001 ry=0 rz=-1.4195 rad; joints [-73.886, -68.929, -104.178, -96.885, 90.142, -82.58] deg
            SuppressedNode
              Set DigitalOutput pin=digital_out[5]; digitalValue=1
            SuppressedNode
              MoveL speed 250 mm/s, acceleration 1200 mm/s^2 (useActiveTCP=true optimoveEnabled=false optiMoveSpeed=0.3 optiMoveAcceleration=0.09) feature=Base
                Waypoint Waypoint_22: motionParameters(jointSpeed=1.047198 jointAcceleration=1.396263 cartesianSpeed=0.1 cartesianAcceleration=0.5); TCP in base x=-31.771 y=-348.512 z=220.918 mm, rx=0.0001 ry=0 rz=-1.1964 rad; joints [-72.82, -67.691, -123.366, -78.936, 90.15, -94.217] deg
                Waypoint Waypoint_23: motionParameters(jointSpeed=1.047198 jointAcceleration=1.396263 cartesianSpeed=0.05 cartesianAcceleration=0.3); TCP in base x=-31.891 y=-348.193 z=178.714 mm, rx=0.0001 ry=0 rz=-1.1964 rad; joints [-72.841, -69.405, -128.724, -71.864, 90.145, -94.213] deg
            SuppressedNode
              Set DigitalOutput pin=digital_out[5]; digitalValue=0
            SuppressedNode
              Wait Sleep waitTime=1
            SuppressedNode
              URCap Gripper (Robotiq_Grippers, Robotiq Inc.) dataModel(position=0.0, force=30.19607843137255, speed=40.0, positionInDouble=0.0, forceInDouble=30.19607843137255, speedInDouble=40.0, slaveIds=[9], blocking=true)
            SuppressedNode
              MoveL speed 250 mm/s, acceleration 1200 mm/s^2 (useActiveTCP=true optimoveEnabled=false optiMoveSpeed=0.3 optiMoveAcceleration=0.09) feature=Base
                Waypoint Waypoint_24: motionParameters(jointSpeed=1.047198 jointAcceleration=1.396263 cartesianSpeed=0.05 cartesianAcceleration=0.3); TCP in base x=-31.773 y=-348.52 z=270.997 mm, rx=0.0001 ry=0 rz=-1.1964 rad; joints [-72.799, -66.725, -116.549, -86.72, 90.151, -94.226] deg
            SuppressedNode
              SafeHome (positionOptionType=SPEED_AND_ACCELERATION speed=1.047198 acceleration=1.396263 nextMotionTime=2)
      SuppressedNode
        Case (caseValue=36)
          SuppressedNode
            MoveL speed 250 mm/s, acceleration 1200 mm/s^2 (useActiveTCP=true optimoveEnabled=false optiMoveSpeed=0.3 optiMoveAcceleration=0.09) feature=Base
              Waypoint Waypoint_26: TCP in base x=-30.182 y=-347.336 z=210.998 mm, rx=0 ry=0 rz=0 rad; joints [-72.486, -67.792, -124.787, -77.413, 90.141, -162.427] deg
          SuppressedNode
            URCap Gripper (Robotiq_Grippers, Robotiq Inc.) dataModel(position=100.0, force=30.19607843137255, speed=40.0, positionInDouble=100.0, forceInDouble=30.19607843137255, speedInDouble=40.0, slaveIds=[9], blocking=true)
          SuppressedNode
            Folder Decap
              Action_Info := "decapping"
              Set DigitalOutput pin=GRP_3F_Enable; digitalValue=1
              Set DigitalOutput pin=GRP_3F_Decap; digitalValue=1
              Force Frame feature=Base; selection=[0, 0, 1, 0, 0, 0]; wrench=[0, 0, 1, 0, 0, 0]; limitsForce=[0.15, 0.15, 0.001, 1.047198, 1.047198, 1.047198]; limitsMotion=[0.1, 0.1, 0.1, 0.349066, 0.349066, 0.349066]
                Script: check_decapping(offset=0.015, timeout=12, abort=CMD_Hold)
              Set DigitalOutput pin=GRP_3F_Decap; digitalValue=0
              Set DigitalOutput pin=GRP_3F_Enable; digitalValue=0
              MoveL speed 250 mm/s, acceleration 1200 mm/s^2 (useActiveTCP=true optimoveEnabled=false optiMoveSpeed=0.3 optiMoveAcceleration=0.09) feature=Base
                Waypoint Waypoint_27: motionParameters(jointSpeed=1.047198 jointAcceleration=1.396263 cartesianSpeed=0.1 cartesianAcceleration=0.5 blendRadius=0.05); TCP in base x=-30.361 y=-347.415 z=279.539 mm, rx=0 ry=0 rz=-0.0004 rad; joints [-72.488, -66.465, -115.449, -88.079, 90.139, -162.449] deg
                Waypoint Waypoint_28: motionParameters(jointSpeed=1.047198 jointAcceleration=1.396263 cartesianSpeed=0.1 cartesianAcceleration=0.5 blendRadius=0.05); TCP in base x=-154.725 y=-473.257 z=246.189 mm, rx=0 ry=0 rz=-0.0004 rad; joints [-92.526, -89.454, -102.579, -77.959, 90.132, -182.495] deg
                Waypoint Waypoint_29: motionParameters(jointSpeed=1.047198 jointAcceleration=1.396263 cartesianSpeed=0.1 cartesianAcceleration=0.3); TCP in base x=-145.695 y=-485.909 z=46.677 mm, rx=0 ry=0 rz=-0.0004 rad; joints [-91.444, -104.036, -119.144, -46.812, 90.094, -181.324] deg
              URCap Gripper (Robotiq_Grippers, Robotiq Inc.) dataModel(position=61.24306326304106, force=30.19607843137255, speed=40.0, positionInDouble=61.24306326304106, forceInDouble=30.19607843137255, speedInDouble=40.0, slaveIds=[9], blocking=true)
              MoveL speed 250 mm/s, acceleration 1200 mm/s^2 (useActiveTCP=true optimoveEnabled=false optiMoveSpeed=0.3 optiMoveAcceleration=0.09) feature=Base
                Waypoint Waypoint_38: motionParameters(jointSpeed=1.047198 jointAcceleration=1.396263 cartesianSpeed=0.1 cartesianAcceleration=0.5 blendRadius=0.05); TCP in base x=-145.695 y=-485.909 z=261.43 mm, rx=0 ry=0 rz=-0.0004 rad; joints [-91.4, -90.37, -99.399, -80.223, 90.132, -181.38] deg
                URCap Gripper (Robotiq_Grippers, Robotiq Inc.) dataModel(position=0.0, force=30.19607843137255, speed=40.0, positionInDouble=0.0, forceInDouble=30.19607843137255, speedInDouble=40.0, slaveIds=[9], blocking=true)
                Waypoint Waypoint_30: motionParameters(jointSpeed=1.047198 jointAcceleration=1.396263 cartesianSpeed=0.1 cartesianAcceleration=0.5 blendRadius=0.05); TCP in base x=-30.182 y=-347.336 z=265.578 mm, rx=0 ry=0 rz=0 rad; joints [-72.462, -66.558, -117.437, -85.997, 90.142, -162.436] deg
                Waypoint Waypoint_31: motionParameters(jointSpeed=1.047198 jointAcceleration=1.396263 cartesianSpeed=0.1 cartesianAcceleration=0.5); TCP in base x=-30.182 y=-347.336 z=175.833 mm, rx=0 ry=0 rz=0 rad; joints [-72.5, -69.38, -129.182, -71.43, 90.136, -162.42] deg
              URCap Gripper (Robotiq_Grippers, Robotiq Inc.) dataModel(position=79.44506104328524, force=30.19607843137255, speed=40.0, positionInDouble=79.44506104328524, forceInDouble=30.19607843137255, speedInDouble=40.0, slaveIds=[9], blocking=true)
              Wait Sleep waitTime=1
              Set DigitalOutput pin=digital_out[5]; digitalValue=1
              MoveL speed 250 mm/s, acceleration 1200 mm/s^2 (useActiveTCP=true optimoveEnabled=false optiMoveSpeed=0.3 optiMoveAcceleration=0.09) feature=Base
                Waypoint Waypoint_32: motionParameters(jointSpeed=1.047198 jointAcceleration=1.396263 cartesianSpeed=0.1 cartesianAcceleration=0.5 blendRadius=0.05); TCP in base x=-30.182 y=-347.336 z=316.067 mm, rx=0 ry=0 rz=0 rad; joints [-72.438, -66.521, -110.081, -93.39, 90.138, -162.442] deg
              URCap VISOR Robotic App (SensoPart VISOR Robotic, SensoPart Industriesensorik GmbH) dataModel(visorAppTemplate=1); state(isChildrenLocked=true)
                URCap Easy Pick Setup (SensoPart VISOR Robotic, SensoPart Industriesensorik GmbH) dataModel(visorId=0, visorSetJob=true, visorJobName=Weigh_scale, visorImageAcqSetup=2, visorImageAcqSource=1, visorCalibSetNo=9, visorDetector=1, visorSetupStatus=5, visorOffsetSet=true, Pose(key=visorGripPose, Position(key=posePosition, Length(key=X value=-0.66092 unit=M), Length(key=Y value=-0.026261 unit=M), Length(key=Z value=0.113423 unit=M)), Rotation(key=poseRotation, Angle(key=RX value=0.044036 unit=RAD), Angle(key=RY value=-0.006733 unit=RAD), Angle(key=RZ value=-1.658906 unit=RAD)))); state(isChildrenLocked=true)
                URCap Process (SensoPart VISOR Robotic, SensoPart Industriesensorik GmbH) dataModel(Variable(key=visorCounterVar, variable=easyPickCount_2), Variable(key=visorPartsFoundVar, variable=easyPickParts_2)); state(isChildrenLocked=true)
                  URCap Image Acquisition Pose (SensoPart VISOR Robotic, SensoPart Industriesensorik GmbH) state(isChildrenLocked=true)
                  URCap Object Detected (SensoPart VISOR Robotic, SensoPart Industriesensorik GmbH) state(isChildrenLocked=true)
                    Folder Open Gripper
                      Wait NoWait
                    URCap Approach Pose (SensoPart VISOR Robotic, SensoPart Industriesensorik GmbH) dataModel(visorOffsetZ=-50.0); state(isChildrenLocked=true)
                    URCap Target Pose (SensoPart VISOR Robotic, SensoPart Industriesensorik GmbH) state(isChildrenLocked=true)
                    Folder Close Gripper
                      URCap Gripper (Robotiq_Grippers, Robotiq Inc.) dataModel(position=0.0, force=30.19607843137255, speed=40.0, positionInDouble=0.0, forceInDouble=30.19607843137255, speedInDouble=40.0, slaveIds=[9], blocking=true)
                    URCap Exit Pose (SensoPart VISOR Robotic, SensoPart Industriesensorik GmbH) dataModel(visorOffsetZ=-100.0); state(isChildrenLocked=true)
                  URCap No Object Detected (SensoPart VISOR Robotic, SensoPart Industriesensorik GmbH) dataModel(Variable(key=visorNoObjCountVar, variable=easyPickNoObj_2))
                    Popup Message (haltProgram=false message=No weigh scale is detected inputType=Text)
              SafeHome (positionOptionType=SPEED_AND_ACCELERATION speed=1.047198 acceleration=1.396263 nextMotionTime=2)
              MoveJ speed 60 deg/s, acceleration 80 deg/s^2 (useActiveTCP=true optimoveEnabled=false optiMoveSpeed=0.3 optiMoveAcceleration=0.09) feature=Base
                Waypoint Waypoint_39: TCP in base x=137.772 y=-577.76 z=300 mm, rx=0 ry=0 rz=-1.5944 rad; joints [-63.54, -101.785, -81.001, -87.198, 90.144, -62.245] deg
              MoveL speed 250 mm/s, acceleration 1200 mm/s^2 (useActiveTCP=true optimoveEnabled=false optiMoveSpeed=0.3 optiMoveAcceleration=0.09) feature=Base
                Waypoint Waypoint_41: motionParameters(jointSpeed=1.047198 jointAcceleration=1.396263 cartesianSpeed=0.1 cartesianAcceleration=0.5); TCP in base x=74.223 y=-565.642 z=234.62 mm, rx=-0.5169 ry=0.5292 rz=-1.5296 rad; joints [-54.985, -107.527, -85.329, -102.066, 60.279, -46.981] deg
                Waypoint Waypoint_40: motionParameters(jointSpeed=1.047198 jointAcceleration=1.396263 cartesianSpeed=0.05 cartesianAcceleration=0.3); TCP in base x=39.988 y=-564.833 z=191.055 mm, rx=-0.7676 ry=0.3431 rz=-2.2413 rad; joints [-57.701, -107.406, -92.471, -93.607, 59.17, -6.639] deg
              URCap Gripper (Robotiq_Grippers, Robotiq Inc.) dataModel(position=100.0, force=20.0, speed=30.0, positionInDouble=100.0, forceInDouble=20.0, speedInDouble=30.0, slaveIds=[9], blocking=true)
              Loop Counting (count=2) loopVariable=Loop_2
                MoveL speed 250 mm/s, acceleration 1200 mm/s^2 (useActiveTCP=true optimoveEnabled=false optiMoveSpeed=0.3 optiMoveAcceleration=0.09) feature=Base
                  Waypoint Waypoint_42: motionParameters(jointSpeed=1.047198 jointAcceleration=1.396263 cartesianSpeed=0.5 cartesianAcceleration=1.2 blendRadius=0); TCP in base x=41.363 y=-564.865 z=192.806 mm, rx=0.2785 ry=0.6241 rz=0.7623 rad; joints [-57.586, -107.397, -92.198, -93.963, 59.209, -186.442] deg
                  Waypoint Waypoint_43: TCP in base x=41.363 y=-564.865 z=192.806 mm, rx=0.9734 ry=0.0641 rz=2.8083 rad; joints [-57.585, -107.391, -92.207, -93.949, 59.207, -310.817] deg
                URCap Gripper (Robotiq_Grippers, Robotiq Inc.) dataModel(position=24.83906770255271, force=20.0, speed=30.19607843137255, positionInDouble=24.83906770255271, forceInDouble=20.0, speedInDouble=30.19607843137255, slaveIds=[9], blocking=true)
                MoveL speed 250 mm/s, acceleration 1200 mm/s^2 (useActiveTCP=true optimoveEnabled=false optiMoveSpeed=0.3 optiMoveAcceleration=0.09) feature=Base
                  Waypoint Waypoint_44: motionParameters(jointSpeed=1.047198 jointAcceleration=1.396263 cartesianSpeed=0.5 cartesianAcceleration=1.2 blendRadius=0); TCP in base x=40.883 y=-564.854 z=192.194 mm, rx=0.1109 ry=0.6592 rz=0.2757 rad; joints [-57.626, -107.402, -92.291, -93.842, 59.196, -157.494] deg
                  Waypoint Waypoint_45: TCP in base x=42.648 y=-564.896 z=194.439 mm, rx=-0.4517 ry=0.5632 rz=-1.3434 rad; joints [-57.484, -107.381, -91.951, -94.273, 59.256, -60.779] deg
                URCap Gripper (Robotiq_Grippers, Robotiq Inc.) dataModel(position=78.43137254901961, force=20.0, speed=30.0, positionInDouble=78.43137254901961, forceInDouble=20.0, speedInDouble=30.0, slaveIds=[9], blocking=true)
              MoveL speed 250 mm/s, acceleration 1200 mm/s^2 (useActiveTCP=true optimoveEnabled=false optiMoveSpeed=0.3 optiMoveAcceleration=0.09) feature=Base
                Waypoint Waypoint_46: motionParameters(jointSpeed=1.047198 jointAcceleration=1.396263 cartesianSpeed=0.05 cartesianAcceleration=0.3); TCP in base x=99.944 y=-566.244 z=267.343 mm, rx=-0.4517 ry=0.5632 rz=-1.3434 rad; joints [-53.041, -108.287, -79.23, -108.385, 61.102, -56.184] deg
                Waypoint Waypoint_47: motionParameters(jointSpeed=1.047198 jointAcceleration=1.396263 cartesianSpeed=0.1 cartesianAcceleration=0.5 blendRadius=0); TCP in base x=99.944 y=-566.244 z=267.343 mm, rx=-0.1017 ry=0.0587 rz=-1.4579 rad; joints [-63.671, -99.121, -88.981, -82.751, 84.056, -70.038] deg
                Waypoint Waypoint_48: motionParameters(jointSpeed=1.047198 jointAcceleration=1.396263 cartesianSpeed=0.25 cartesianAcceleration=1.2); TCP in base x=-136.183 y=-647.487 z=294.248 mm, rx=-0.1017 ry=0.0587 rz=-1.4579 rad; joints [-87.788, -109.526, -72.49, -86.263, 84.243, -94.331] deg
                Waypoint Waypoint_49: TCP in base x=-159.024 y=-641.021 z=47.692 mm, rx=0 ry=0 rz=-1.4579 rad; joints [-92.238, -121.266, -92.571, -56.15, 90.14, -98.675] deg
              URCap Gripper (Robotiq_Grippers, Robotiq Inc.) dataModel(position=33.9400665926748, force=20.0, speed=30.19607843137255, positionInDouble=33.9400665926748, forceInDouble=20.0, speedInDouble=30.19607843137255, slaveIds=[9], blocking=true)
              MoveL speed 250 mm/s, acceleration 1200 mm/s^2 (useActiveTCP=true optimoveEnabled=false optiMoveSpeed=0.3 optiMoveAcceleration=0.09) feature=Base
                Waypoint Waypoint_50: TCP in base x=-159.024 y=-641.021 z=291.114 mm, rx=0 ry=0 rz=-1.4579 rad; joints [-92.2, -111.308, -69.838, -88.841, 90.151, -98.75] deg
                SafeHome (positionOptionType=SPEED_AND_ACCELERATION speed=1.047198 acceleration=1.396263 nextMotionTime=2)
      SuppressedNode
        Case (caseValue=37)
          SuppressedNode
            URCap VISOR Robotic App (SensoPart VISOR Robotic, SensoPart Industriesensorik GmbH) dataModel(visorAppTemplate=1); state(isChildrenLocked=true)
              URCap Easy Pick Setup (SensoPart VISOR Robotic, SensoPart Industriesensorik GmbH) dataModel(visorId=0, visorSetJob=true, visorJobName=Spatula, visorImageAcqSetup=2, visorImageAcqSource=1, visorCalibSetNo=10, visorDetector=1, visorOffsetSet=true, visorSetupStatus=5, Pose(key=visorGripPose, Position(key=posePosition, Length(key=X value=-0.64401 unit=M), Length(key=Y value=-0.309906 unit=M), Length(key=Z value=0.133972 unit=M)), Rotation(key=poseRotation, Angle(key=RX value=0.000082 unit=RAD), Angle(key=RY value=0.000005 unit=RAD), Angle(key=RZ value=3.001273 unit=RAD)))); state(isChildrenLocked=true)
              URCap Process (SensoPart VISOR Robotic, SensoPart Industriesensorik GmbH) dataModel(Variable(key=visorCounterVar, variable=easyPickCount_3), Variable(key=visorPartsFoundVar, variable=easyPickParts_3)); state(isChildrenLocked=true)
                URCap Image Acquisition Pose (SensoPart VISOR Robotic, SensoPart Industriesensorik GmbH) state(isChildrenLocked=true)
                URCap Object Detected (SensoPart VISOR Robotic, SensoPart Industriesensorik GmbH) state(isChildrenLocked=true)
                  Folder Open Gripper
                    URCap Gripper (Robotiq_Grippers, Robotiq Inc.) dataModel(position=0.0, force=20.0, speed=30.19607843137255, positionInDouble=0.0, forceInDouble=20.0, speedInDouble=30.19607843137255, slaveIds=[9], blocking=true)
                  URCap Approach Pose (SensoPart VISOR Robotic, SensoPart Industriesensorik GmbH) dataModel(visorOffsetZ=-100.0); state(isChildrenLocked=true)
                  URCap Target Pose (SensoPart VISOR Robotic, SensoPart Industriesensorik GmbH) state(isChildrenLocked=true)
                  Folder Close Gripper
                    URCap Gripper (Robotiq_Grippers, Robotiq Inc.) dataModel(position=100.0, force=20.0, speed=30.19607843137255, positionInDouble=100.0, forceInDouble=20.0, speedInDouble=30.19607843137255, slaveIds=[9], blocking=true)
                  URCap Exit Pose (SensoPart VISOR Robotic, SensoPart Industriesensorik GmbH) dataModel(visorToolSpeed=100.0, visorToolAcc=300.0, visorOffsetZ=-200.0); state(isChildrenLocked=true)
                URCap No Object Detected (SensoPart VISOR Robotic, SensoPart Industriesensorik GmbH) dataModel(Variable(key=visorNoObjCountVar, variable=easyPickNoObj_3))
                  Popup Message (haltProgram=false message=No spatula is detected inputType=Text)
          URCap VISOR Robotic App (SensoPart VISOR Robotic, SensoPart Industriesensorik GmbH) dataModel(visorAppTemplate=1); state(isChildrenLocked=true)
            URCap Easy Pick Setup (SensoPart VISOR Robotic, SensoPart Industriesensorik GmbH) dataModel(visorId=0, visorSetJob=true, visorJobName=Spatula_horizontal, visorImageAcqSetup=2, visorImageAcqSource=0, visorDetector=1, visorOffsetSet=true, visorSetupStatus=1, Pose(key=visorImageAcqPose, Position(key=posePosition, Length(key=X value=-0.477866 unit=M), Length(key=Y value=0.377208 unit=M), Length(key=Z value=0.48314 unit=M)), Rotation(key=poseRotation, Angle(key=RX value=-0.000072 unit=RAD), Angle(key=RY value=-0.000033 unit=RAD), Angle(key=RZ value=-1.610249 unit=RAD))), Pose(key=visorGripPose, Position(key=posePosition, Length(key=X value=-0.547139 unit=M), Length(key=Y value=0.33515 unit=M), Length(key=Z value=0.041533 unit=M)), Rotation(key=poseRotation, Angle(key=RX value=2.188123 unit=RAD), Angle(key=RY value=-0.020843 unit=RAD), Angle(key=RZ value=2.219811 unit=RAD)))); state(isChildrenLocked=true)
            URCap Process (SensoPart VISOR Robotic, SensoPart Industriesensorik GmbH) dataModel(Variable(key=visorCounterVar, variable=easyPickCount_5), Variable(key=visorPartsFoundVar, variable=easyPickParts_5)); state(isChildrenLocked=true)
              URCap Image Acquisition Pose (SensoPart VISOR Robotic, SensoPart Industriesensorik GmbH) state(isChildrenLocked=true)
              URCap Object Detected (SensoPart VISOR Robotic, SensoPart Industriesensorik GmbH) state(isChildrenLocked=true)
                Folder Open Gripper
                  URCap Gripper (Robotiq_Grippers, Robotiq Inc.) dataModel(position=43.04106548279689, force=30.0, speed=30.0, positionInDouble=43.04106548279689, forceInDouble=30.0, speedInDouble=30.0, slaveIds=[9], blocking=true)
                URCap Approach Pose (SensoPart VISOR Robotic, SensoPart Industriesensorik GmbH) dataModel(visorOffsetZ=-130.0); state(isChildrenLocked=true)
                URCap Target Pose (SensoPart VISOR Robotic, SensoPart Industriesensorik GmbH) state(isChildrenLocked=true)
                Folder Close Gripper
                  URCap Gripper (Robotiq_Grippers, Robotiq Inc.) dataModel(position=100.0, force=30.0, speed=30.0, positionInDouble=100.0, forceInDouble=30.0, speedInDouble=30.0, slaveIds=[9], blocking=true)
                URCap Exit Pose (SensoPart VISOR Robotic, SensoPart Industriesensorik GmbH) dataModel(visorOffsetZ=-170.0); state(isChildrenLocked=true)
              URCap No Object Detected (SensoPart VISOR Robotic, SensoPart Industriesensorik GmbH) dataModel(Variable(key=visorNoObjCountVar, variable=easyPickNoObj_5))
                Popup Message (haltProgram=false message=No Spatula detected inputType=Text)
          SuppressedNode
            MoveJ speed 60 deg/s, acceleration 80 deg/s^2 (useActiveTCP=true optimoveEnabled=false optiMoveSpeed=0.3 optiMoveAcceleration=0.09) feature=Base
              Waypoint Waypoint_1: motionParameters(jointSpeed=1.047198 jointAcceleration=1.396263 cartesianSpeed=0.1 cartesianAcceleration=0.5 blendRadius=0.05); TCP in base x=-359.544 y=319.273 z=259.271 mm, rx=2.1553 ry=-0.0199 rz=2.2443 rad; joints [-228.189, -86.975, -126.838, -149.463, 223.669, -271.634] deg
              Waypoint Waypoint_51: motionParameters(jointSpeed=1.047198 jointAcceleration=1.396263 cartesianSpeed=0.1 cartesianAcceleration=0.5 blendRadius=0); TCP in base x=-477.866 y=377.208 z=483.14 mm, rx=-0.0001 ry=0 rz=-1.6102 rad; joints [-205.499, -110.086, -42.439, -117.467, 90.106, -203.428] deg
              Waypoint Waypoint_52: TCP in base x=-42.31 y=-356.333 z=399.894 mm, rx=0 ry=0 rz=-0.1228 rad; joints [-74.871, -69.823, -95.716, -104.453, 90.124, -157.892] deg
          MoveL speed 50 mm/s, acceleration 300 mm/s^2 (useActiveTCP=true optimoveEnabled=false optiMoveSpeed=0.3 optiMoveAcceleration=0.09) feature=Base
            Waypoint Waypoint_3: motionParameters(jointSpeed=1.047198 jointAcceleration=1.396263 cartesianSpeed=0.05 cartesianAcceleration=0.3); TCP in base x=-31.864 y=-349.975 z=230.259 mm, rx=0 ry=0 rz=0 rad; joints [-72.901, -67.669, -121.993, -80.33, 90.142, -162.853] deg
            Waypoint Waypoint_80: motionParameters(jointSpeed=1.047198 jointAcceleration=1.396263 cartesianSpeed=0.05 cartesianAcceleration=0.3); TCP in base x=143.03 y=-569.853 z=275.754 mm, rx=1.2979 ry=0.0264 rz=2.7129 rad; joints [-47.784, -117.454, -67.716, -126.008, 56.917, 63.329] deg
            Loop Counting (count=3) loopVariable=Loop_3
              Waypoint Waypoint_55: motionParameters(jointSpeed=1.047198 jointAcceleration=1.396263 cartesianSpeed=0.05 cartesianAcceleration=0.3); TCP in base x=73.857 y=-577.013 z=221.505 mm, rx=1.2979 ry=0.0264 rz=2.7129 rad; joints [-52.913, -114.774, -80.289, -113.397, 53.656, 58.584] deg
                Until TOOL_CONTACT_DETECTION (allowActions=false retraction=0 decelerationAcceleration=3 decelerationAngularAcceleration=34.906585)
              Waypoint Waypoint_56: motionParameters(jointSpeed=1.047198 jointAcceleration=1.396263 cartesianSpeed=0.05 cartesianAcceleration=0.3); TCP in base x=135.677 y=-579.448 z=242.231 mm, rx=1.5554 ry=0.0154 rz=2.5559 rad; joints [-47.427, -124.812, -65.265, -134.284, 52.841, 72.036] deg
            Loop Counting (count=2) loopVariable=Loop_5
              Waypoint Waypoint_56: motionParameters(jointSpeed=1.047198 jointAcceleration=1.396263 cartesianSpeed=0.05 cartesianAcceleration=0.3); TCP in base x=135.677 y=-579.448 z=242.231 mm, rx=1.5554 ry=0.0154 rz=2.5559 rad; joints [-47.427, -124.812, -65.265, -134.284, 52.841, 72.036] deg
              Waypoint Waypoint_101: motionParameters(jointSpeed=1.047198 jointAcceleration=1.396263 cartesianSpeed=0.5 cartesianAcceleration=1.2); TCP in base x=143.391 y=-581.809 z=226.065 mm, rx=1.6397 ry=0.0079 rz=2.5024 rad; joints [-46.773, -128.399, -63.349, -137.511, 52.317, 75.293] deg
            Waypoint Waypoint_59: motionParameters(jointSpeed=1.047198 jointAcceleration=1.396263 cartesianSpeed=0.05 cartesianAcceleration=0.3); TCP in base x=272.401 y=-578.183 z=239.561 mm, rx=2.127 ry=0.1139 rz=2.1556 rad; joints [-37.816, -154.733, -25.502, -178.522, 53.445, 96.624] deg
            Waypoint Waypoint_58: motionParameters(jointSpeed=1.047198 jointAcceleration=1.396263 cartesianSpeed=0.05 cartesianAcceleration=0.3); TCP in base x=223.649 y=-578.478 z=276.546 mm, rx=2.1743 ry=-0.0441 rz=2.0587 rad; joints [-41.771, -153.265, -25.455, -184.54, 55.381, 96.631] deg
          MoveJ speed 30 deg/s, acceleration 50 deg/s^2 (useActiveTCP=true optimoveEnabled=false optiMoveSpeed=0.3 optiMoveAcceleration=0.09) feature=Base
            Waypoint Waypoint_60: motionParameters(jointSpeed=0.349066 jointAcceleration=0.523599 cartesianSpeed=0.25 cartesianAcceleration=1.2 blendRadius=0.05); TCP in base x=-13.316 y=-544.772 z=383.372 mm, rx=2.2082 ry=0.0375 rz=2.0976 rad; joints [-53.447, -120.321, -68.514, -175.377, 39.556, 98.101] deg
            Waypoint Waypoint_61: motionParameters(jointSpeed=0.349066 jointAcceleration=0.523599 cartesianSpeed=0.25 cartesianAcceleration=1.2 blendRadius=0.05); TCP in base x=-412.189 y=-356.447 z=383.372 mm, rx=1.7517 ry=-0.74 rz=1.6007 rad; joints [-101.195, -120.321, -68.514, -175.377, 39.556, 98.101] deg
            Waypoint Waypoint_62: motionParameters(jointSpeed=0.349066 jointAcceleration=0.523599 cartesianSpeed=0.25 cartesianAcceleration=1.2); TCP in base x=-542.659 y=-114.282 z=251.262 mm, rx=1.813 ry=-0.6794 rz=1.6553 rad; joints [-123.661, -111.262, -103.952, -159.22, 12.548, 108.767] deg
          MoveL speed 250 mm/s, acceleration 1200 mm/s^2 (useActiveTCP=true optimoveEnabled=false optiMoveSpeed=0.3 optiMoveAcceleration=0.09) feature=Base
            Waypoint Waypoint_63: motionParameters(jointSpeed=1.047198 jointAcceleration=1.396263 cartesianSpeed=0.05 cartesianAcceleration=0.3); TCP in base x=-532.496 y=-127.81 z=159.342 mm, rx=1.813 ry=-0.6794 rz=1.6553 rad; joints [-121.654, -119.526, -108.357, -144.665, 14.532, 106.823] deg
            Waypoint Waypoint_102: motionParameters(jointSpeed=1.047198 jointAcceleration=1.396263 cartesianSpeed=0.05 cartesianAcceleration=0.3); TCP in base x=-576.035 y=-66.27 z=306.74 mm, rx=0.8621 ry=-0.2554 rz=2.1952 rad; joints [-142.141, -87.685, -107.535, -64.498, 50.077, -8.596] deg
            Waypoint Waypoint_103: motionParameters(jointSpeed=1.047198 jointAcceleration=1.396263 cartesianSpeed=0.05 cartesianAcceleration=0.3); TCP in base x=-581.965 y=-59.291 z=312.082 mm, rx=0.8621 ry=-0.2554 rz=2.1952 rad; joints [-143.275, -88.018, -106.65, -64.116, 50.29, -10.05] deg
            Waypoint Waypoint_81: motionParameters(jointSpeed=1.047198 jointAcceleration=1.396263 cartesianSpeed=0.5 cartesianAcceleration=1.2); TCP in base x=-581.965 y=-59.291 z=290.576 mm, rx=0.8621 ry=-0.2554 rz=2.1952 rad; joints [-143.281, -88.87, -109.094, -60.824, 50.286, -10.043] deg
            Waypoint Decap_above: TCP in base x=-31.864 y=-349.975 z=288.042 mm, rx=0 ry=0 rz=0 rad; joints [-72.875, -66.865, -113.978, -89.149, 90.141, -162.862] deg
          MoveJ speed 60 deg/s, acceleration 80 deg/s^2 (useActiveTCP=true optimoveEnabled=false optiMoveSpeed=0.3 optiMoveAcceleration=0.09) feature=Base
            Waypoint Waypoint_104: TCP in base x=-333.293 y=-480.744 z=350.142 mm, rx=2.2175 ry=0.1409 rz=2.2091 rad; joints [-82.414, -101.687, -97.87, -162.913, 4.302, 96.426] deg
          SuppressedNode
            Weight_value := get_weight()
      SuppressedNode
        Case (caseValue=38)
          SuppressedNode
            URCap VISOR Robotic App (SensoPart VISOR Robotic, SensoPart Industriesensorik GmbH) dataModel(visorAppTemplate=1); state(isChildrenLocked=true)
              URCap Easy Pick Setup (SensoPart VISOR Robotic, SensoPart Industriesensorik GmbH) dataModel(visorId=0, visorSetJob=true, visorJobName=Container_S_rack, visorImageAcqSetup=2, visorSetupStatus=2); state(isChildrenLocked=true)
              URCap Process (SensoPart VISOR Robotic, SensoPart Industriesensorik GmbH) dataModel(Variable(key=visorCounterVar, variable=easyPickCount_4), Variable(key=visorPartsFoundVar, variable=easyPickParts_4)); state(isChildrenLocked=true)
                URCap Image Acquisition Pose (SensoPart VISOR Robotic, SensoPart Industriesensorik GmbH) state(isChildrenLocked=true)
                URCap Object Detected (SensoPart VISOR Robotic, SensoPart Industriesensorik GmbH) state(isChildrenLocked=true)
                  Folder Open Gripper
                    Placeholder
                  URCap Approach Pose (SensoPart VISOR Robotic, SensoPart Industriesensorik GmbH) state(isChildrenLocked=true)
                  URCap Target Pose (SensoPart VISOR Robotic, SensoPart Industriesensorik GmbH) state(isChildrenLocked=true)
                  Folder Close Gripper
                    Placeholder
                  URCap Exit Pose (SensoPart VISOR Robotic, SensoPart Industriesensorik GmbH) state(isChildrenLocked=true)
                URCap No Object Detected (SensoPart VISOR Robotic, SensoPart Industriesensorik GmbH) dataModel(Variable(key=visorNoObjCountVar, variable=easyPickNoObj_4))
                  Placeholder
      Case (caseValue=39)
        Folder Powder container Pick [hidden by the author, left out]
      Case (caseValue=40)
        Folder Decap Container  [hidden by the author, left out]
      Case (caseValue=41)
        Folder Place the open PowderA container & dosing
          SuppressedNode
            Script: tilt_to_home()
          SuppressedNode
            Script: tilt_send(4)
          URCap VISOR Robotic App (SensoPart VISOR Robotic, SensoPart Industriesensorik GmbH) dataModel(visorAppTemplate=1); state(isChildrenLocked=true)
            URCap Easy Pick Setup (SensoPart VISOR Robotic, SensoPart Industriesensorik GmbH) dataModel(visorId=0, visorImageAcqSetup=2, visorDetector=1, visorSetJob=true, visorOffsetSet=true, visorImageAcqSource=2, visorJobName=PoTS, visorSetupStatus=4, Pose(key=visorGripPose, Position(key=posePosition, Length(key=X value=-0.726236 unit=M), Length(key=Y value=-0.14014 unit=M), Length(key=Z value=0.266183 unit=M)), Rotation(key=poseRotation, Angle(key=RX value=-0.811878 unit=RAD), Angle(key=RY value=1.689668 unit=RAD), Angle(key=RZ value=-1.713453 unit=RAD))), Feature(key=visorImageAcqFeature name=Trigger)); state(isChildrenLocked=true)
            URCap Process (SensoPart VISOR Robotic, SensoPart Industriesensorik GmbH) dataModel(Variable(key=visorCounterVar, variable=easyPickCount_7), Variable(key=visorPartsFoundVar, variable=easyPickParts_7)); state(isChildrenLocked=true)
              URCap Image Acquisition Pose (SensoPart VISOR Robotic, SensoPart Industriesensorik GmbH) state(isChildrenLocked=true)
              URCap Object Detected (SensoPart VISOR Robotic, SensoPart Industriesensorik GmbH) state(isChildrenLocked=true)
                Folder Open Gripper
                  URCap Gripper (Robotiq_Grippers, Robotiq Inc.) dataModel(position=0.0, force=30.19607843137255, speed=30.19607843137255, positionInDouble=0.0, forceInDouble=30.19607843137255, speedInDouble=30.19607843137255, slaveIds=[9], blocking=true)
                  MoveL speed 250 mm/s, acceleration 1200 mm/s^2 (useActiveTCP=true optimoveEnabled=false optiMoveSpeed=0.3 optiMoveAcceleration=0.09) feature=Base
                    Waypoint OP_PowderA2: TCP in base x=9.371 y=-409.434 z=294.169 mm, rx=-0.8233 ry=1.7094 rz=-1.6983 rad; joints [-57.265, -122.586, -76.992, -161.25, 72.295, 1.124] deg; TCP offset x=0 y=0 z=161 mm, rx=3.1415 ry=0 rz=0 rad
                    Waypoint OP_PowderA_abov: TCP in base x=-12.145 y=-363.335 z=315.326 mm, rx=-0.7771 ry=1.753 rz=-1.7409 rad; joints [-58.232, -116.012, -83.989, -160.83, 75.01, 1.147] deg; TCP offset x=0 y=0 z=161 mm, rx=3.1415 ry=0 rz=0 rad
                    Waypoint OP_PowderA_pick: TCP in base x=-19.99 y=-367.909 z=180.101 mm, rx=-0.5462 ry=1.936 rz=-1.9301 rad; joints [-66.516, -128.259, -85.768, -146.461, 83.267, 1.188] deg
                    URCap Gripper (Robotiq_Grippers, Robotiq Inc.) dataModel(position=100.0, force=30.19607843137255, speed=30.19607843137255, positionInDouble=100.0, forceInDouble=30.19607843137255, speedInDouble=30.19607843137255, slaveIds=[9], blocking=true)
                    Wait Sleep waitTime=0.5
                    Set DigitalOutput pin=GRP_3F_Open; digitalValue=1
                    SuppressedNode
                      Script: Motors_off()
                    Waypoint OP_PowderA_abov: motionParameters(jointSpeed=1.047198 jointAcceleration=1.396263 cartesianSpeed=0.05 cartesianAcceleration=0.3); TCP in base x=-12.145 y=-363.335 z=315.326 mm, rx=-0.7771 ry=1.753 rz=-1.7409 rad; joints [-58.232, -116.012, -83.989, -160.83, 75.01, 1.147] deg
                    Waypoint Op_PowA_wP: TCP in base x=-173.728 y=-372.934 z=295.117 mm, rx=-0.9724 ry=1.541 rz=-1.5487 rad; joints [-67.269, -106.894, -99.849, -153.52, 49.211, 1.028] deg
                URCap Approach Pose (SensoPart VISOR Robotic, SensoPart Industriesensorik GmbH) dataModel(visorOffsetZ=0.0, visorJointSpeed=25.0, visorJointAcc=30.0); state(isChildrenLocked=true)
                URCap Target Pose (SensoPart VISOR Robotic, SensoPart Industriesensorik GmbH) dataModel(visorToolSpeed=50.0, visorToolAcc=100.0); state(isChildrenLocked=true)
                Folder Close Gripper
                  container_place := get_actual_tcp_pose()
                  target_pose := pose_add(container_place, p[0,0,-0.1,0,0,0])
                  MoveL speed 250 mm/s, acceleration 1200 mm/s^2 (useActiveTCP=true optimoveEnabled=false optiMoveSpeed=0.3 optiMoveAcceleration=0.09) feature=Base
                    Waypoint Variable (Variable): motionParameters(jointSpeed=1.047198 jointAcceleration=1.396263 cartesianSpeed=0.05 cartesianAcceleration=0.3); variable=target_pose
                  URCap Gripper (Robotiq_Grippers, Robotiq Inc.) dataModel(position=0.0, force=30.19607843137255, speed=30.19607843137255, positionInDouble=0.0, forceInDouble=30.19607843137255, speedInDouble=30.19607843137255, slaveIds=[9], blocking=true)
                URCap Exit Pose (SensoPart VISOR Robotic, SensoPart Industriesensorik GmbH) dataModel(visorOffsetZ=0.0); state(isChildrenLocked=true)
              URCap No Object Detected (SensoPart VISOR Robotic, SensoPart Industriesensorik GmbH) dataModel(Variable(key=visorNoObjCountVar, variable=easyPickNoObj_7))
                Popup Message (haltProgram=false message=No weigh scale detected inputType=Text)
          place_pose := get_actual_tcp_pose()
          Script: center_pose()
          SuppressedNode
            center_tilt_pos := P_center
          MoveJ speed 60 deg/s, acceleration 80 deg/s^2 (useActiveTCP=true optimoveEnabled=false optiMoveSpeed=0.3 optiMoveAcceleration=0.09) feature=Base
            Waypoint Waypoint_1: TCP in base x=-451.049 y=-340.589 z=308.224 mm, rx=0.0971 ry=0.091 rz=-1.5784 rad; joints [-127.334, -100.578, -80.109, -94.907, 86.186, -126.663] deg
      Case (caseValue=42)
        Folder Powder Emptying [hidden by the author, left out]
      Case (caseValue=43)
        Folder Powder dosing
          SuppressedNode
            Script: zero_scale()
          Script: send_target_info()
          Script: send_powder_info()
          SuppressedNode
            Folder spatula_selection test
              weight_value := get_weight()
              diff := target_weight-weight_value
              Script: scooping_init()
              Script: compute_level_percent(W_now, weight_value)
              Script: spatula = select_spatula(Pow_name, level, diff)
          URCap VISOR Robotic App (SensoPart VISOR Robotic, SensoPart Industriesensorik GmbH) dataModel(visorAppTemplate=1); state(isChildrenLocked=true)
            URCap Easy Pick Setup (SensoPart VISOR Robotic, SensoPart Industriesensorik GmbH) dataModel(visorId=0, visorSetJob=true, visorImageAcqSetup=2, visorCalibSetNo=9, visorDetector=1, visorImageAcqSource=2, visorJobName=Weight_scale, visorOffsetSet=true, visorSetupStatus=3, Pose(key=visorGripPose, Position(key=posePosition, Length(key=X value=-0.535221 unit=M), Length(key=Y value=0.017694 unit=M), Length(key=Z value=0.123958 unit=M)), Rotation(key=poseRotation, Angle(key=RX value=0.727814 unit=RAD), Angle(key=RY value=1.465761 unit=RAD), Angle(key=RZ value=-0.763944 unit=RAD))), Feature(key=visorImageAcqFeature name=Trigger)); state(isChildrenLocked=true)
            URCap Process (SensoPart VISOR Robotic, SensoPart Industriesensorik GmbH) dataModel(Variable(key=visorCounterVar, variable=easyPickCount_4), Variable(key=visorPartsFoundVar, variable=easyPickParts_4)); state(isChildrenLocked=true)
              URCap Image Acquisition Pose (SensoPart VISOR Robotic, SensoPart Industriesensorik GmbH) state(isChildrenLocked=true)
              URCap Object Detected (SensoPart VISOR Robotic, SensoPart Industriesensorik GmbH) state(isChildrenLocked=true)
                Folder Open Gripper
                  Script: tare_scale()
                  Wait Sleep waitTime=0.2
                  weight_value := get_weight()
                  Wait Sleep waitTime=0.2
                  diff := target_weight-weight_value
                  Script: scooping_init()
                  Script: compute_level_percent(W_now, weight_value)
                  Script: send_level_info()
                  Script: spatula = select_spatula(Pow_name, level, diff)
                  Wait Sleep waitTime=0.2
                  Script: send_spatula_info()
                  If spatula ≟ "spatula_L"
                    MoveJ speed 60 deg/s, acceleration 80 deg/s^2 (useActiveTCP=true optimoveEnabled=false optiMoveSpeed=0.3 optiMoveAcceleration=0.09) feature=Base
                      Waypoint Spatula_otw: TCP in base x=-38.472 y=-263.141 z=425.351 mm, rx=-0.0004 ry=-0.0001 rz=3.0344 rad; joints [-68.119, -57.773, -97.702, -114.504, 90.127, 27.957] deg
                      Waypoint pick_spat_L_abv: TCP in base x=239.059 y=-67.213 z=280.721 mm, rx=0 ry=-0.0005 rz=3.1068 rad; joints [16.774, -49.077, -122.624, -98.282, 90.162, 108.776] deg
                    MoveL speed 250 mm/s, acceleration 1200 mm/s^2 (useActiveTCP=true optimoveEnabled=false optiMoveSpeed=0.3 optiMoveAcceleration=0.09) feature=Base
                      Waypoint spat_L_pick: TCP in base x=242.469 y=-67.302 z=193.171 mm, rx=0 ry=-0.0005 rz=3.1068 rad; joints [16.429, -49.275, -135.385, -85.324, 90.17, 108.483] deg
                      URCap Gripper (Robotiq_Grippers, Robotiq Inc.) dataModel(position=100.0, force=30.0, speed=0.0, positionInDouble=100.0, forceInDouble=30.0, speedInDouble=0.0, slaveIds=[9], blocking=true)
                      Waypoint spat_L_lift: motionParameters(blendRadius=0.01); TCP in base x=245.402 y=-67.432 z=289.049 mm, rx=0 ry=-0.0005 rz=3.1068 rad; joints [16.24, -50.411, -121.005, -98.568, 90.16, 108.238] deg
                      Waypoint spat_L_side: motionParameters(blendRadius=0.01); TCP in base x=247.134 y=-17.634 z=289.063 mm, rx=0 ry=-0.0005 rz=3.1068 rad; joints [28.487, -49.174, -121.365, -99.443, 90.16, 120.484] deg
